  movel([-0.251057, -0.840337, -2.769867, -1.102185, 1.570796, 1.319739],accel_mss,speed_ms,0,blend_radius_m)
  movel([-0.250306, -0.839240, -2.770084, -1.103065, 1.570796, 1.320491],accel_mss,speed_ms,0,blend_radius_m)
  movel([-0.248421, -0.837227, -2.770480, -1.104681, 1.570796, 1.322375],accel_mss,speed_ms,0,blend_radius_m)
  movel([-0.247261, -0.836341, -2.770654, -1.105394, 1.570796, 1.323536],accel_mss,speed_ms,0,blend_radius_m)
  movel([-0.246051, -0.835788, -2.770763, -1.105839, 1.570796, 1.324746],accel_mss,speed_ms,0,blend_radius_m)
  movel([-0.245067, -0.835822, -2.770756, -1.105811, 1.570796, 1.325730],accel_mss,speed_ms,0,blend_radius_m)
  movel([-0.243698, -0.836942, -2.770537, -1.104911, 1.570796, 1.327098],accel_mss,speed_ms,0,blend_radius_m)
  movel([-0.242450, -0.839139, -2.770104, -1.103146, 1.570796, 1.328347],accel_mss,speed_ms,0,blend_radius_m)
  movel([-0.241508, -0.841625, -2.769611, -1.101153, 1.570796, 1.329288],accel_mss,speed_ms,0,blend_radius_m)
  movel([-0.239706, -0.837507, -2.770425, -1.104456, 1.570796, 1.331091],accel_mss,speed_ms,0,blend_radius_m)
  movel([-0.237551, -0.833302, -2.771247, -1.107840, 1.570796, 1.333246],accel_mss,speed_ms,0,blend_radius_m)
  movel([-0.235089, -0.829066, -2.772064, -1.111259, 1.570796, 1.335707],accel_mss,speed_ms,0,blend_radius_m)
  movel([-0.232380, -0.824862, -2.772866, -1.114661, 1.570796, 1.338416],accel_mss,speed_ms,0,blend_radius_m)
  movel([-0.226936, -0.816422, -2.774445, -1.121522, 1.570796, 1.343860],accel_mss,speed_ms,0,blend_radius_m)
  movel([-0.225279, -0.814079, -2.774877, -1.123434, 1.570796, 1.345517],accel_mss,speed_ms,0,blend_radius_m)
  movel([-0.223613, -0.811962, -2.775264, -1.125163, 1.570796, 1.347184],accel_mss,speed_ms,0,blend_radius_m)
  movel([-0.221984, -0.810225, -2.775580, -1.126584, 1.570796, 1.348813],accel_mss,speed_ms,0,blend_radius_m)
  movel([-0.220457, -0.809030, -2.775796, -1.127562, 1.570796, 1.350339],accel_mss,speed_ms,0,blend_radius_m)
  movel([-0.219063, -0.808558, -2.775882, -1.127949, 1.570796, 1.351734],accel_mss,speed_ms,0,blend_radius_m)
  movel([-0.217966, -0.808858, -2.775828, -1.127704, 1.570796, 1.352830],accel_mss,speed_ms,0,blend_radius_m)
  movel([-0.217165, -0.809769, -2.775663, -1.126958, 1.570796, 1.353632],accel_mss,speed_ms,0,blend_radius_m)
  movel([-0.216671, -0.811136, -2.775414, -1.125838, 1.570796, 1.354126],accel_mss,speed_ms,0,blend_radius_m)
  movel([-0.216485, -0.812799, -2.775111, -1.124479, 1.570796, 1.354311],accel_mss,speed_ms,0,blend_radius_m)
  movel([-0.216608, -0.814592, -2.774782, -1.123014, 1.570796, 1.354188],accel_mss,speed_ms,0,blend_radius_m)
  movel([-0.217044, -0.816361, -2.774456, -1.121571, 1.570796, 1.353752],accel_mss,speed_ms,0,blend_radius_m)
  movel([-0.217800, -0.817948, -2.774162, -1.120278, 1.570796, 1.352996],accel_mss,speed_ms,0,blend_radius_m)
  movel([-0.212688, -0.810429, -2.775543, -1.126417, 1.570796, 1.358108],accel_mss,speed_ms,0,blend_radius_m)
  movel([-0.209894, -0.806731, -2.776211, -1.129447, 1.570796, 1.360902],accel_mss,speed_ms,0,blend_radius_m)
  movel([-0.206949, -0.803115, -2.776856, -1.132417, 1.570796, 1.363847],accel_mss,speed_ms,0,blend_radius_m)
  movel([-0.203868, -0.799614, -2.777475, -1.135300, 1.570796, 1.366928],accel_mss,speed_ms,0,blend_radius_m)
  movel([-0.200656, -0.796258, -2.778062, -1.138069, 1.570796, 1.370141],accel_mss,speed_ms,0,blend_radius_m)
  movel([-0.197322, -0.793081, -2.778612, -1.140696, 1.570796, 1.373474],accel_mss,speed_ms,0,blend_radius_m)
  movel([-0.193879, -0.790113, -2.779121, -1.143155, 1.570796, 1.376917],accel_mss,speed_ms,0,blend_radius_m)
  movel([-0.191467, -0.788517, -2.779393, -1.144480, 1.570796, 1.379330],accel_mss,speed_ms,0,blend_radius_m)
  movel([-0.188786, -0.787373, -2.779587, -1.145430, 1.570796, 1.382010],accel_mss,speed_ms,0,blend_radius_m)
  movel([-0.187580, -0.787128, -2.779628, -1.145633, 1.570796, 1.383216],accel_mss,speed_ms,0,blend_radius_m)
  movel([-0.186584, -0.787179, -2.779619, -1.145591, 1.570796, 1.384213],accel_mss,speed_ms,0,blend_radius_m)
  movel([-0.185886, -0.787588, -2.779550, -1.145251, 1.570796, 1.384910],accel_mss,speed_ms,0,blend_radius_m)
  movel([-0.185586, -0.788421, -2.779409, -1.144559, 1.570796, 1.385210],accel_mss,speed_ms,0,blend_radius_m)
  movel([-0.185771, -0.789581, -2.779211, -1.143597, 1.570796, 1.385025],accel_mss,speed_ms,0,blend_radius_m)
  movel([-0.186325, -0.790924, -2.778982, -1.142483, 1.570796, 1.384471],accel_mss,speed_ms,0,blend_radius_m)
  movel([-0.188126, -0.794006, -2.778452, -1.139931, 1.570796, 1.382670],accel_mss,speed_ms,0,blend_radius_m)
  movel([-0.190402, -0.796962, -2.777939, -1.137488, 1.570796, 1.380394],accel_mss,speed_ms,0,blend_radius_m)
  movel([-0.192970, -0.799746, -2.777452, -1.135191, 1.570796, 1.377827],accel_mss,speed_ms,0,blend_radius_m)
  movel([-0.195646, -0.802312, -2.776999, -1.133078, 1.570796, 1.375151],accel_mss,speed_ms,0,blend_radius_m)
  movel([-0.191927, -0.800596, -2.777302, -1.134491, 1.570796, 1.378869],accel_mss,speed_ms,0,blend_radius_m)
  movel([-0.188109, -0.798487, -2.777673, -1.136229, 1.570796, 1.382688],accel_mss,speed_ms,0,blend_radius_m)
  movel([-0.184228, -0.796012, -2.778104, -1.138273, 1.570796, 1.386568],accel_mss,speed_ms,0,blend_radius_m)
  movel([-0.180320, -0.793191, -2.778593, -1.140606, 1.570796, 1.390476],accel_mss,speed_ms,0,blend_radius_m)
  movel([-0.177275, -0.790678, -2.779024, -1.142687, 1.570796, 1.393522],accel_mss,speed_ms,0,blend_radius_m)
  movel([-0.171365, -0.785323, -2.779933, -1.147134, 1.570796, 1.399431],accel_mss,speed_ms,0,blend_radius_m)
  movel([-0.168296, -0.782767, -2.780361, -1.149261, 1.570796, 1.402501],accel_mss,speed_ms,0,blend_radius_m)
  movel([-0.164758, -0.780078, -2.780808, -1.151503, 1.570796, 1.406038],accel_mss,speed_ms,0,blend_radius_m)
  movel([-0.158752, -0.775824, -2.781507, -1.155058, 1.570796, 1.412044],accel_mss,speed_ms,0,blend_radius_m)
  movel([-0.155841, -0.774007, -2.781803, -1.156579, 1.570796, 1.414955],accel_mss,speed_ms,0,blend_radius_m)
  movel([-0.153543, -0.772881, -2.781986, -1.157523, 1.570796, 1.417254],accel_mss,speed_ms,0,blend_radius_m)
  movel([-0.152751, -0.772687, -2.782017, -1.157685, 1.570796, 1.418046],accel_mss,speed_ms,0,blend_radius_m)
  movel([-0.152271, -0.772806, -2.781998, -1.157586, 1.570796, 1.418525],accel_mss,speed_ms,0,blend_radius_m)
  movel([-0.152148, -0.773270, -2.781923, -1.157196, 1.570796, 1.418648],accel_mss,speed_ms,0,blend_radius_m)
  movel([-0.152440, -0.774130, -2.781783, -1.156476, 1.570796, 1.418357],accel_mss,speed_ms,0,blend_radius_m)
  movel([-0.153723, -0.776356, -2.781420, -1.154613, 1.570796, 1.417074],accel_mss,speed_ms,0,blend_radius_m)
  movel([-0.155470, -0.778742, -2.781028, -1.152619, 1.570796, 1.415326],accel_mss,speed_ms,0,blend_radius_m)
  movel([-0.157553, -0.781219, -2.780619, -1.150552, 1.570796, 1.413244],accel_mss,speed_ms,0,blend_radius_m)
  movel([-0.159834, -0.783698, -2.780205, -1.148485, 1.570796, 1.410962],accel_mss,speed_ms,0,blend_radius_m)
  movel([-0.164497, -0.788374, -2.779417, -1.144598, 1.570796, 1.406299],accel_mss,speed_ms,0,blend_radius_m)
  movel([-0.168438, -0.792159, -2.778770, -1.141460, 1.570796, 1.402358],accel_mss,speed_ms,0,blend_radius_m)
  movel([-0.166238, -0.791550, -2.778875, -1.141964, 1.570796, 1.404559],accel_mss,speed_ms,0,blend_radius_m)
  movel([-0.163950, -0.790704, -2.779020, -1.142666, 1.570796, 1.406846],accel_mss,speed_ms,0,blend_radius_m)
  movel([-0.159176, -0.788425, -2.779408, -1.144556, 1.570796, 1.411620],accel_mss,speed_ms,0,blend_radius_m)
  movel([-0.154224, -0.785549, -2.779894, -1.146946, 1.570796, 1.416572],accel_mss,speed_ms,0,blend_radius_m)
  movel([-0.149200, -0.782306, -2.780438, -1.149645, 1.570796, 1.421597],accel_mss,speed_ms,0,blend_radius_m)
  movel([-0.145052, -0.779396, -2.780920, -1.152073, 1.570796, 1.425744],accel_mss,speed_ms,0,blend_radius_m)
  movel([-0.132523, -0.770152, -2.782425, -1.159811, 1.570796, 1.438273],accel_mss,speed_ms,0,blend_radius_m)
  movel([-0.130147, -0.768779, -2.782645, -1.160965, 1.570796, 1.440650],accel_mss,speed_ms,0,blend_radius_m)
  movel([-0.128213, -0.768174, -2.782742, -1.161473, 1.570796, 1.442583],accel_mss,speed_ms,0,blend_radius_m)
  movel([-0.127762, -0.768378, -2.782709, -1.161302, 1.570796, 1.443034],accel_mss,speed_ms,0,blend_radius_m)
  movel([-0.127842, -0.769035, -2.782604, -1.160750, 1.570796, 1.442955],accel_mss,speed_ms,0,blend_radius_m)
  movel([-0.128593, -0.770230, -2.782413, -1.159746, 1.570796, 1.442203],accel_mss,speed_ms,0,blend_radius_m)
  movel([-0.130154, -0.772048, -2.782120, -1.158221, 1.570796, 1.440642],accel_mss,speed_ms,0,blend_radius_m)
  movel([-0.132825, -0.774737, -2.781684, -1.155968, 1.570796, 1.437971],accel_mss,speed_ms,0,blend_radius_m)
  movel([-0.135952, -0.777548, -2.781225, -1.153616, 1.570796, 1.434844],accel_mss,speed_ms,0,blend_radius_m)
  movel([-0.139084, -0.779981, -2.780824, -1.151585, 1.570796, 1.431712],accel_mss,speed_ms,0,blend_radius_m)
  movel([-0.140515, -0.780901, -2.780671, -1.150816, 1.570796, 1.430281],accel_mss,speed_ms,0,blend_radius_m)
  movel([-0.141777, -0.781533, -2.780566, -1.150290, 1.570796, 1.429020],accel_mss,speed_ms,0,blend_radius_m)
  movel([-0.136604, -0.780701, -2.780705, -1.150984, 1.570796, 1.434192],accel_mss,speed_ms,0,blend_radius_m)
  movel([-0.131148, -0.779248, -2.780945, -1.152196, 1.570796, 1.439648],accel_mss,speed_ms,0,blend_radius_m)
  movel([-0.125468, -0.777292, -2.781267, -1.153830, 1.570796, 1.445329],accel_mss,speed_ms,0,blend_radius_m)
  movel([-0.119612, -0.774952, -2.781649, -1.155788, 1.570796, 1.451185],accel_mss,speed_ms,0,blend_radius_m)
  movel([-0.107622, -0.769590, -2.782515, -1.160284, 1.570796, 1.463175],accel_mss,speed_ms,0,blend_radius_m)
  movel([-0.095682, -0.764142, -2.783380, -1.164866, 1.570796, 1.475114],accel_mss,speed_ms,0,blend_radius_m)
  movel([-0.093660, -0.763518, -2.783479, -1.165393, 1.570796, 1.477136],accel_mss,speed_ms,0,blend_radius_m)
  movel([-0.092947, -0.763655, -2.783457, -1.165277, 1.570796, 1.477849],accel_mss,speed_ms,0,blend_radius_m)
  movel([-0.092662, -0.764296, -2.783356, -1.164736, 1.570796, 1.478134],accel_mss,speed_ms,0,blend_radius_m)
  movel([-0.092897, -0.765328, -2.783193, -1.163868, 1.570796, 1.477899],accel_mss,speed_ms,0,blend_radius_m)
  movel([-0.094551, -0.768317, -2.782719, -1.161353, 1.570796, 1.476245],accel_mss,speed_ms,0,blend_radius_m)
  movel([-0.095791, -0.770072, -2.782438, -1.159879, 1.570796, 1.475005],accel_mss,speed_ms,0,blend_radius_m)
  movel([-0.098671, -0.773409, -2.781900, -1.157080, 1.570796, 1.472125],accel_mss,speed_ms,0,blend_radius_m)
  movel([-0.101929, -0.776471, -2.781401, -1.154516, 1.570796, 1.468867],accel_mss,speed_ms,0,blend_radius_m)
  movel([-0.105410, -0.779237, -2.780947, -1.152206, 1.570796, 1.465387],accel_mss,speed_ms,0,blend_radius_m)
  movel([-0.108946, -0.781663, -2.780545, -1.150181, 1.570796, 1.461850],accel_mss,speed_ms,0,blend_radius_m)
  movel([-0.112381, -0.783724, -2.780201, -1.148464, 1.570796, 1.458416],accel_mss,speed_ms,0,blend_radius_m)
  movel([-0.115557, -0.785382, -2.779923, -1.147085, 1.570796, 1.455240],accel_mss,speed_ms,0,blend_radius_m)
  movel([-0.118308, -0.786594, -2.779718, -1.146077, 1.570796, 1.452489],accel_mss,speed_ms,0,blend_radius_m)
  movel([-0.118229, -0.787293, -2.779600, -1.145496, 1.570796, 1.452568],accel_mss,speed_ms,0,blend_radius_m)
  movel([-0.117672, -0.787561, -2.779555, -1.145274, 1.570796, 1.453124],accel_mss,speed_ms,0,blend_radius_m)
  movel([-0.116060, -0.787683, -2.779534, -1.145172, 1.570796, 1.454736],accel_mss,speed_ms,0,blend_radius_m)
  movel([-0.114280, -0.787508, -2.779564, -1.145318, 1.570796, 1.456517],accel_mss,speed_ms,0,blend_radius_m)
  movel([-0.110443, -0.786631, -2.779712, -1.146046, 1.570796, 1.460353],accel_mss,speed_ms,0,blend_radius_m)
  movel([-0.103651, -0.784713, -2.780035, -1.147641, 1.570796, 1.467145],accel_mss,speed_ms,0,blend_radius_m)
  movel([-0.096773, -0.782536, -2.780399, -1.149454, 1.570796, 1.474024],accel_mss,speed_ms,0,blend_radius_m)
  movel([-0.082734, -0.777500, -2.781233, -1.153657, 1.570796, 1.488063],accel_mss,speed_ms,0,blend_radius_m)
  movel([-0.078824, -0.776168, -2.781451, -1.154770, 1.570796, 1.491972],accel_mss,speed_ms,0,blend_radius_m)
  movel([-0.076323, -0.775517, -2.781557, -1.155315, 1.570796, 1.494474],accel_mss,speed_ms,0,blend_radius_m)
  movel([-0.073893, -0.775133, -2.781620, -1.155636, 1.570796, 1.496903],accel_mss,speed_ms,0,blend_radius_m)
  movel([-0.071878, -0.775218, -2.781606, -1.155565, 1.570796, 1.498918],accel_mss,speed_ms,0,blend_radius_m)
  movel([-0.070612, -0.775956, -2.781486, -1.154948, 1.570796, 1.500184],accel_mss,speed_ms,0,blend_radius_m)
  movel([-0.070357, -0.776623, -2.781377, -1.154390, 1.570796, 1.500439],accel_mss,speed_ms,0,blend_radius_m)
  movel([-0.070410, -0.777522, -2.781229, -1.153638, 1.570796, 1.500387],accel_mss,speed_ms,0,blend_radius_m)
  movel([-0.070817, -0.778683, -2.781038, -1.152668, 1.570796, 1.499979],accel_mss,speed_ms,0,blend_radius_m)
  movel([-0.071609, -0.780115, -2.780802, -1.151472, 1.570796, 1.499188],accel_mss,speed_ms,0,blend_radius_m)
  movel([-0.072883, -0.781500, -2.780572, -1.150317, 1.570796, 1.497913],accel_mss,speed_ms,0,blend_radius_m)
  movel([-0.074697, -0.782890, -2.780340, -1.149159, 1.570796, 1.496099],accel_mss,speed_ms,0,blend_radius_m)
  movel([-0.084551, -0.789376, -2.779246, -1.143767, 1.570796, 1.486245],accel_mss,speed_ms,0,blend_radius_m)
  movel([-0.087910, -0.791177, -2.778939, -1.142274, 1.570796, 1.482886],accel_mss,speed_ms,0,blend_radius_m)
  movel([-0.089384, -0.791747, -2.778841, -1.141801, 1.570796, 1.481412],accel_mss,speed_ms,0,blend_radius_m)
  movel([-0.090634, -0.791996, -2.778798, -1.141595, 1.570796, 1.480162],accel_mss,speed_ms,0,blend_radius_m)
  movel([-0.085187, -0.792592, -2.778696, -1.141101, 1.570796, 1.485610],accel_mss,speed_ms,0,blend_radius_m)
  movel([-0.079266, -0.792365, -2.778735, -1.141289, 1.570796, 1.491530],accel_mss,speed_ms,0,blend_radius_m)
  movel([-0.072987, -0.791466, -2.778889, -1.142034, 1.570796, 1.497810],accel_mss,speed_ms,0,blend_radius_m)
  movel([-0.066459, -0.790039, -2.779133, -1.143217, 1.570796, 1.504338],accel_mss,speed_ms,0,blend_radius_m)
  movel([-0.060916, -0.788133, -2.779458, -1.144799, 1.570796, 1.509880],accel_mss,speed_ms,0,blend_radius_m)
  movel([-0.052946, -0.785532, -2.779897, -1.146959, 1.570796, 1.517850],accel_mss,speed_ms,0,blend_radius_m)
  movel([-0.049278, -0.784724, -2.780033, -1.147631, 1.570796, 1.521518],accel_mss,speed_ms,0,blend_radius_m)
  movel([-0.046471, -0.784631, -2.780049, -1.147709, 1.570796, 1.524326],accel_mss,speed_ms,0,blend_radius_m)
  movel([-0.045545, -0.784943, -2.779996, -1.147450, 1.570796, 1.525252],accel_mss,speed_ms,0,blend_radius_m)
  movel([-0.045021, -0.785541, -2.779896, -1.146953, 1.570796, 1.525776],accel_mss,speed_ms,0,blend_radius_m)
  movel([-0.044956, -0.786463, -2.779740, -1.146186, 1.570796, 1.525840],accel_mss,speed_ms,0,blend_radius_m)
  movel([-0.045403, -0.787732, -2.779526, -1.145131, 1.570796, 1.525393],accel_mss,speed_ms,0,blend_radius_m)
  movel([-0.046180, -0.789074, -2.779298, -1.144017, 1.570796, 1.524616],accel_mss,speed_ms,0,blend_radius_m)
  movel([-0.047117, -0.790379, -2.779075, -1.142935, 1.570796, 1.523680],accel_mss,speed_ms,0,blend_radius_m)
  movel([-0.049250, -0.792857, -2.778650, -1.140882, 1.570796, 1.521546],accel_mss,speed_ms,0,blend_radius_m)
  movel([-0.051649, -0.795339, -2.778221, -1.138829, 1.570796, 1.519147],accel_mss,speed_ms,0,blend_radius_m)
  movel([-0.056596, -0.799831, -2.777437, -1.135121, 1.570796, 1.514200],accel_mss,speed_ms,0,blend_radius_m)
  movel([-0.059113, -0.801820, -2.777086, -1.133483, 1.570796, 1.511683],accel_mss,speed_ms,0,blend_radius_m)
  movel([-0.054139, -0.800667, -2.777290, -1.134433, 1.570796, 1.516658],accel_mss,speed_ms,0,blend_radius_m)
  movel([-0.049049, -0.799176, -2.777552, -1.135662, 1.570796, 1.521747],accel_mss,speed_ms,0,blend_radius_m)
  movel([-0.043853, -0.797385, -2.777865, -1.137138, 1.570796, 1.526944],accel_mss,speed_ms,0,blend_radius_m)
  movel([-0.038557, -0.795324, -2.778224, -1.138841, 1.570796, 1.532239],accel_mss,speed_ms,0,blend_radius_m)
  movel([-0.027716, -0.790540, -2.779048, -1.142802, 1.570796, 1.543080],accel_mss,speed_ms,0,blend_radius_m)
  movel([-0.016601, -0.785088, -2.779972, -1.147329, 1.570796, 1.554196],accel_mss,speed_ms,0,blend_radius_m)
  movel([-0.013645, -0.783918, -2.780168, -1.148302, 1.570796, 1.557151],accel_mss,speed_ms,0,blend_radius_m)
  movel([-0.012527, -0.783932, -2.780166, -1.148291, 1.570796, 1.558270],accel_mss,speed_ms,0,blend_radius_m)
  movel([-0.011960, -0.784664, -2.780043, -1.147681, 1.570796, 1.558836],accel_mss,speed_ms,0,blend_radius_m)
  movel([-0.011973, -0.785494, -2.779904, -1.146991, 1.570796, 1.558823],accel_mss,speed_ms,0,blend_radius_m)
  movel([-0.012257, -0.786461, -2.779741, -1.146187, 1.570796, 1.558540],accel_mss,speed_ms,0,blend_radius_m)
  movel([-0.013515, -0.788743, -2.779354, -1.144292, 1.570796, 1.557281],accel_mss,speed_ms,0,blend_radius_m)
  movel([-0.015472, -0.791310, -2.778916, -1.142163, 1.570796, 1.555324],accel_mss,speed_ms,0,blend_radius_m)
  movel([-0.017868, -0.793984, -2.778456, -1.139949, 1.570796, 1.552928],accel_mss,speed_ms,0,blend_radius_m)
  movel([-0.022942, -0.798903, -2.777600, -1.135886, 1.570796, 1.547854],accel_mss,speed_ms,0,blend_radius_m)
  movel([-0.026708, -0.802032, -2.777048, -1.133308, 1.570796, 1.544089],accel_mss,speed_ms,0,blend_radius_m)
  movel([-0.024456, -0.801160, -2.777202, -1.134026, 1.570796, 1.546340],accel_mss,speed_ms,0,blend_radius_m)
  movel([-0.022148, -0.800059, -2.777397, -1.134934, 1.570796, 1.548648],accel_mss,speed_ms,0,blend_radius_m)
  movel([-0.017405, -0.797244, -2.777890, -1.137255, 1.570796, 1.553391],accel_mss,speed_ms,0,blend_radius_m)
  movel([-0.012565, -0.793690, -2.778507, -1.140192, 1.570796, 1.558232],accel_mss,speed_ms,0,blend_radius_m)
  movel([-0.007710, -0.789520, -2.779222, -1.143648, 1.570796, 1.563087],accel_mss,speed_ms,0,blend_radius_m)
  movel([-0.002926, -0.784828, -2.780016, -1.147546, 1.570796, 1.567870],accel_mss,speed_ms,0,blend_radius_m)
  movel([0.001697, -0.779740, -2.780864, -1.151785, 1.570796, 1.572493],accel_mss,speed_ms,0,blend_radius_m)
  movel([0.006066, -0.774361, -2.781746, -1.156282, 1.570796, 1.576863],accel_mss,speed_ms,0,blend_radius_m)
  movel([0.010091, -0.768815, -2.782639, -1.160935, 1.570796, 1.580887],accel_mss,speed_ms,0,blend_radius_m)
  movel([0.011867, -0.766339, -2.783033, -1.163017, 1.570796, 1.582663],accel_mss,speed_ms,0,blend_radius_m)
  movel([0.012853, -0.765231, -2.783209, -1.163949, 1.570796, 1.583649],accel_mss,speed_ms,0,blend_radius_m)
  movel([0.013911, -0.764336, -2.783350, -1.164703, 1.570796, 1.584707],accel_mss,speed_ms,0,blend_radius_m)
  movel([0.015047, -0.763769, -2.783439, -1.165181, 1.570796, 1.585844],accel_mss,speed_ms,0,blend_radius_m)
  movel([0.016045, -0.763599, -2.783466, -1.165324, 1.570796, 1.586842],accel_mss,speed_ms,0,blend_radius_m)
  movel([0.017197, -0.764007, -2.783402, -1.164980, 1.570796, 1.587993],accel_mss,speed_ms,0,blend_radius_m)
  movel([0.017895, -0.765128, -2.783225, -1.164036, 1.570796, 1.588691],accel_mss,speed_ms,0,blend_radius_m)
  movel([0.018210, -0.766786, -2.782962, -1.162640, 1.570796, 1.589006],accel_mss,speed_ms,0,blend_radius_m)
  movel([0.018221, -0.768822, -2.782638, -1.160929, 1.570796, 1.589018],accel_mss,speed_ms,0,blend_radius_m)
  movel([0.017618, -0.773331, -2.781913, -1.157145, 1.570796, 1.588414],accel_mss,speed_ms,0,blend_radius_m)
  movel([0.016685, -0.777318, -2.781263, -1.153808, 1.570796, 1.587481],accel_mss,speed_ms,0,blend_radius_m)
  movel([0.020069, -0.771975, -2.782132, -1.158282, 1.570796, 1.590865],accel_mss,speed_ms,0,blend_radius_m)
  movel([0.023040, -0.766596, -2.782993, -1.162801, 1.570796, 1.593836],accel_mss,speed_ms,0,blend_radius_m)
  movel([0.025578, -0.761235, -2.783836, -1.167318, 1.570796, 1.596375],accel_mss,speed_ms,0,blend_radius_m)
  movel([0.027672, -0.755966, -2.784651, -1.171772, 1.570796, 1.598468],accel_mss,speed_ms,0,blend_radius_m)
  movel([0.029286, -0.750858, -2.785427, -1.176104, 1.570796, 1.600082],accel_mss,speed_ms,0,blend_radius_m)
  movel([0.030417, -0.745966, -2.786159, -1.180264, 1.570796, 1.601214],accel_mss,speed_ms,0,blend_radius_m)
  movel([0.031030, -0.741380, -2.786835, -1.184174, 1.570796, 1.601827],accel_mss,speed_ms,0,blend_radius_m)
  movel([0.031110, -0.737161, -2.787447, -1.187781, 1.570796, 1.601906],accel_mss,speed_ms,0,blend_radius_m)
  movel([0.030356, -0.731952, -2.788191, -1.192246, 1.570796, 1.601153],accel_mss,speed_ms,0,blend_radius_m)
  movel([0.030207, -0.729033, -2.788603, -1.194753, 1.570796, 1.601003],accel_mss,speed_ms,0,blend_radius_m)
  movel([0.030375, -0.727506, -2.788816, -1.196066, 1.570796, 1.601171],accel_mss,speed_ms,0,blend_radius_m)
  movel([0.030771, -0.725941, -2.789034, -1.197414, 1.570796, 1.601568],accel_mss,speed_ms,0,blend_radius_m)
  movel([0.031877, -0.723302, -2.789399, -1.199689, 1.570796, 1.602673],accel_mss,speed_ms,0,blend_radius_m)
  movel([0.033028, -0.721615, -2.789630, -1.201144, 1.570796, 1.603824],accel_mss,speed_ms,0,blend_radius_m)
  movel([0.034209, -0.720678, -2.789758, -1.201953, 1.570796, 1.605005],accel_mss,speed_ms,0,blend_radius_m)
  movel([0.035393, -0.720293, -2.789810, -1.202286, 1.570796, 1.606190],accel_mss,speed_ms,0,blend_radius_m)
  movel([0.038713, -0.720456, -2.789788, -1.202145, 1.570796, 1.609509],accel_mss,speed_ms,0,blend_radius_m)
  movel([0.039670, -0.720273, -2.789813, -1.202303, 1.570796, 1.610466],accel_mss,speed_ms,0,blend_radius_m)
  movel([0.041218, -0.716370, -2.790341, -1.205678, 1.570796, 1.612014],accel_mss,speed_ms,0,blend_radius_m)
  movel([0.042449, -0.712549, -2.790850, -1.208990, 1.570796, 1.613245],accel_mss,speed_ms,0,blend_radius_m)
  movel([0.043380, -0.708824, -2.791341, -1.212224, 1.570796, 1.614176],accel_mss,speed_ms,0,blend_radius_m)
  movel([0.044028, -0.705202, -2.791811, -1.215376, 1.570796, 1.614824],accel_mss,speed_ms,0,blend_radius_m)
  movel([0.044398, -0.701705, -2.792260, -1.218424, 1.570796, 1.615194],accel_mss,speed_ms,0,blend_radius_m)
  movel([0.044507, -0.698341, -2.792686, -1.221362, 1.570796, 1.615303],accel_mss,speed_ms,0,blend_radius_m)
  movel([0.044023, -0.692041, -2.793470, -1.226877, 1.570796, 1.614819],accel_mss,speed_ms,0,blend_radius_m)
  movel([0.042690, -0.686413, -2.794156, -1.231820, 1.570796, 1.613487],accel_mss,speed_ms,0,blend_radius_m)
  movel([0.040657, -0.681528, -2.794740, -1.236121, 1.570796, 1.611454],accel_mss,speed_ms,0,blend_radius_m)
  movel([0.038047, -0.677485, -2.795215, -1.239689, 1.570796, 1.608843],accel_mss,speed_ms,0,blend_radius_m)
  movel([0.035023, -0.674343, -2.795579, -1.242467, 1.570796, 1.605819],accel_mss,speed_ms,0,blend_radius_m)
  speed_ms = 0.005
  movel([0.035023, -0.668307, -2.788892, -1.255190, 1.570796, 1.605819],accel_mss,speed_ms,0,blend_radius_m)
  speed_ms = 0.040
  movel([0.005563, -0.693117, -2.785908, -1.233364, 1.570796, 1.576359],accel_mss,speed_ms,0,blend_radius_m)
  speed_ms = 0.005
  movel([0.005563, -0.699497, -2.792540, -1.220352, 1.570796, 1.576359],accel_mss,speed_ms,0,blend_radius_m)
  speed_ms = 0.025
  movel([0.002772, -0.699600, -2.792527, -1.220262, 1.570796, 1.573568],accel_mss,speed_ms,0,blend_radius_m)
  movel([-0.000362, -0.700496, -2.792414, -1.219480, 1.570796, 1.570434],accel_mss,speed_ms,0,blend_radius_m)
  movel([-0.003761, -0.702064, -2.792214, -1.218111, 1.570796, 1.567035],accel_mss,speed_ms,0,blend_radius_m)
  movel([-0.007341, -0.704171, -2.791944, -1.216274, 1.570796, 1.563455],accel_mss,speed_ms,0,blend_radius_m)
  movel([-0.011021, -0.706691, -2.791618, -1.214080, 1.570796, 1.559775],accel_mss,speed_ms,0,blend_radius_m)
  movel([-0.014730, -0.709498, -2.791252, -1.211639, 1.570796, 1.556067],accel_mss,speed_ms,0,blend_radius_m)
  movel([-0.021919, -0.715471, -2.790461, -1.206457, 1.570796, 1.548877],accel_mss,speed_ms,0,blend_radius_m)
  speed_ms = 0.005
  movel([-0.021919, -0.708883, -2.783866, -1.219640, 1.570796, 1.548877],accel_mss,speed_ms,0,blend_radius_m)
  speed_ms = 0.040
  movel([-0.012736, -0.700553, -2.784960, -1.226876, 1.570796, 1.558061],accel_mss,speed_ms,0,blend_radius_m)
  speed_ms = 0.005
  movel([-0.012736, -0.707032, -2.791574, -1.213783, 1.570796, 1.558061],accel_mss,speed_ms,0,blend_radius_m)
  speed_ms = 0.025
  movel([-0.011741, -0.702920, -2.792104, -1.217364, 1.570796, 1.559055],accel_mss,speed_ms,0,blend_radius_m)
  movel([-0.011148, -0.699151, -2.792584, -1.220654, 1.570796, 1.559648],accel_mss,speed_ms,0,blend_radius_m)
  movel([-0.010951, -0.695718, -2.793015, -1.223656, 1.570796, 1.559845],accel_mss,speed_ms,0,blend_radius_m)
  movel([-0.011133, -0.692605, -2.793401, -1.226383, 1.570796, 1.559663],accel_mss,speed_ms,0,blend_radius_m)
  movel([-0.011672, -0.689793, -2.793746, -1.228850, 1.570796, 1.559124],accel_mss,speed_ms,0,blend_radius_m)
  movel([-0.012556, -0.687267, -2.794053, -1.231069, 1.570796, 1.558241],accel_mss,speed_ms,0,blend_radius_m)
  movel([-0.013764, -0.685013, -2.794325, -1.233052, 1.570796, 1.557032],accel_mss,speed_ms,0,blend_radius_m)
  movel([-0.015280, -0.683011, -2.794564, -1.234815, 1.570796, 1.555516],accel_mss,speed_ms,0,blend_radius_m)
  movel([-0.020599, -0.678116, -2.795141, -1.239132, 1.570796, 1.550198],accel_mss,speed_ms,0,blend_radius_m)
  movel([-0.022981, -0.675592, -2.795435, -1.241363, 1.570796, 1.547815],accel_mss,speed_ms,0,blend_radius_m)
  movel([-0.024944, -0.672152, -2.795830, -1.244407, 1.570796, 1.545852],accel_mss,speed_ms,0,blend_radius_m)
  movel([-0.026696, -0.667138, -2.796398, -1.248853, 1.570796, 1.544100],accel_mss,speed_ms,0,blend_radius_m)
  movel([-0.027862, -0.661556, -2.797016, -1.253817, 1.570796, 1.542934],accel_mss,speed_ms,0,blend_radius_m)
  movel([-0.028220, -0.655275, -2.797696, -1.259418, 1.570796, 1.542576],accel_mss,speed_ms,0,blend_radius_m)
  movel([-0.028029, -0.651831, -2.798062, -1.262496, 1.570796, 1.542767],accel_mss,speed_ms,0,blend_radius_m)
  movel([-0.027547, -0.648162, -2.798446, -1.265781, 1.570796, 1.543250],accel_mss,speed_ms,0,blend_radius_m)
  movel([-0.026144, -0.642097, -2.799068, -1.271224, 1.570796, 1.544652],accel_mss,speed_ms,0,blend_radius_m)
  movel([-0.023952, -0.635758, -2.799701, -1.276930, 1.570796, 1.546845],accel_mss,speed_ms,0,blend_radius_m)
  movel([-0.020999, -0.629190, -2.800340, -1.282859, 1.570796, 1.549797],accel_mss,speed_ms,0,blend_radius_m)
  movel([-0.017318, -0.622446, -2.800977, -1.288965, 1.570796, 1.553478],accel_mss,speed_ms,0,blend_radius_m)
  movel([-0.012950, -0.615595, -2.801605, -1.295189, 1.570796, 1.557847],accel_mss,speed_ms,0,blend_radius_m)
  movel([-0.007925, -0.608692, -2.802219, -1.301478, 1.570796, 1.562872],accel_mss,speed_ms,0,blend_radius_m)
  movel([-0.002284, -0.601797, -2.802812, -1.307780, 1.570796, 1.568512],accel_mss,speed_ms,0,blend_radius_m)
  movel([0.003922, -0.594989, -2.803379, -1.314020, 1.570796, 1.574719],accel_mss,speed_ms,0,blend_radius_m)
  movel([0.008850, -0.590063, -2.803778, -1.318548, 1.570796, 1.579646],accel_mss,speed_ms,0,blend_radius_m)
  movel([0.013936, -0.585373, -2.804149, -1.322867, 1.570796, 1.584733],accel_mss,speed_ms,0,blend_radius_m)
  movel([0.019128, -0.580961, -2.804489, -1.326939, 1.570796, 1.589924],accel_mss,speed_ms,0,blend_radius_m)
  movel([0.024383, -0.576845, -2.804800, -1.330743, 1.570796, 1.595179],accel_mss,speed_ms,0,blend_radius_m)
  movel([0.029644, -0.573079, -2.805079, -1.334231, 1.570796, 1.600440],accel_mss,speed_ms,0,blend_radius_m)
  movel([0.034862, -0.569690, -2.805325, -1.337374, 1.570796, 1.605658],accel_mss,speed_ms,0,blend_radius_m)
  movel([0.039979, -0.566716, -2.805537, -1.340135, 1.570796, 1.610775],accel_mss,speed_ms,0,blend_radius_m)
  movel([0.044944, -0.564196, -2.805715, -1.342479, 1.570796, 1.615740],accel_mss,speed_ms,0,blend_radius_m)
  movel([0.049699, -0.562164, -2.805856, -1.344369, 1.570796, 1.620495],accel_mss,speed_ms,0,blend_radius_m)
  movel([0.054199, -0.560647, -2.805960, -1.345782, 1.570796, 1.624995],accel_mss,speed_ms,0,blend_radius_m)
  movel([0.058387, -0.559683, -2.806026, -1.346680, 1.570796, 1.629184],accel_mss,speed_ms,0,blend_radius_m)
  movel([0.062215, -0.559301, -2.806052, -1.347036, 1.570796, 1.633011],accel_mss,speed_ms,0,blend_radius_m)
  movel([0.065633, -0.559525, -2.806036, -1.346827, 1.570796, 1.636430],accel_mss,speed_ms,0,blend_radius_m)
  movel([0.068583, -0.560396, -2.805977, -1.346016, 1.570796, 1.639379],accel_mss,speed_ms,0,blend_radius_m)
  movel([0.071026, -0.561923, -2.805872, -1.344593, 1.570796, 1.641822],accel_mss,speed_ms,0,blend_radius_m)
  movel([0.072920, -0.564138, -2.805719, -1.342532, 1.570796, 1.643716],accel_mss,speed_ms,0,blend_radius_m)
  movel([0.074676, -0.567785, -2.805462, -1.339142, 1.570796, 1.645473],accel_mss,speed_ms,0,blend_radius_m)
  movel([0.075891, -0.571973, -2.805160, -1.335256, 1.570796, 1.646687],accel_mss,speed_ms,0,blend_radius_m)
  movel([0.076668, -0.576581, -2.804820, -1.330988, 1.570796, 1.647464],accel_mss,speed_ms,0,blend_radius_m)
  movel([0.077130, -0.581463, -2.804451, -1.326475, 1.570796, 1.647927],accel_mss,speed_ms,0,blend_radius_m)
  movel([0.077482, -0.592588, -2.803575, -1.316226, 1.570796, 1.648279],accel_mss,speed_ms,0,blend_radius_m)
  movel([0.077191, -0.604219, -2.802606, -1.305564, 1.570796, 1.647987],accel_mss,speed_ms,0,blend_radius_m)
  movel([0.076408, -0.616212, -2.801550, -1.294627, 1.570796, 1.647204],accel_mss,speed_ms,0,blend_radius_m)
  movel([0.075281, -0.628414, -2.800414, -1.283560, 1.570796, 1.646077],accel_mss,speed_ms,0,blend_radius_m)
  movel([0.070103, -0.676768, -2.795298, -1.240323, 1.570796, 1.640899],accel_mss,speed_ms,0,blend_radius_m)
  movel([0.068408, -0.699650, -2.792521, -1.220218, 1.570796, 1.639204],accel_mss,speed_ms,0,blend_radius_m)
  movel([0.067946, -0.710698, -2.791095, -1.210596, 1.570796, 1.638742],accel_mss,speed_ms,0,blend_radius_m)
  movel([0.067855, -0.721372, -2.789663, -1.201354, 1.570796, 1.638651],accel_mss,speed_ms,0,blend_radius_m)
  movel([0.068210, -0.731613, -2.788239, -1.192537, 1.570796, 1.639006],accel_mss,speed_ms,0,blend_radius_m)
  movel([0.069087, -0.741348, -2.786839, -1.184202, 1.570796, 1.639884],accel_mss,speed_ms,0,blend_radius_m)
  movel([0.070552, -0.750526, -2.785477, -1.176385, 1.570796, 1.641348],accel_mss,speed_ms,0,blend_radius_m)
  movel([0.072685, -0.759083, -2.784170, -1.169135, 1.570796, 1.643482],accel_mss,speed_ms,0,blend_radius_m)
  movel([0.073786, -0.762163, -2.783691, -1.166535, 1.570796, 1.644583],accel_mss,speed_ms,0,blend_radius_m)
  movel([0.075340, -0.764775, -2.783281, -1.164333, 1.570796, 1.646136],accel_mss,speed_ms,0,blend_radius_m)
  movel([0.077562, -0.766509, -2.783007, -1.162874, 1.570796, 1.648359],accel_mss,speed_ms,0,blend_radius_m)
  movel([0.078995, -0.766915, -2.782942, -1.162532, 1.570796, 1.649791],accel_mss,speed_ms,0,blend_radius_m)
  movel([0.080684, -0.766942, -2.782938, -1.162510, 1.570796, 1.651480],accel_mss,speed_ms,0,blend_radius_m)
  speed_ms = 0.005
  movel([0.080684, -0.759735, -2.776473, -1.176181, 1.570796, 1.651480],accel_mss,speed_ms,0,blend_radius_m)
  speed_ms = 0.040
  movel([0.042306, -0.732546, -2.780582, -1.199261, 1.570796, 1.613102],accel_mss,speed_ms,0,blend_radius_m)
  speed_ms = 0.005
  movel([0.042306, -0.739433, -2.787118, -1.185838, 1.570796, 1.613102],accel_mss,speed_ms,0,blend_radius_m)
  speed_ms = 0.025
  movel([0.041280, -0.741224, -2.786857, -1.184307, 1.570796, 1.612077],accel_mss,speed_ms,0,blend_radius_m)
  movel([0.040567, -0.743006, -2.786596, -1.182786, 1.570796, 1.611363],accel_mss,speed_ms,0,blend_radius_m)
  movel([0.040141, -0.744758, -2.786338, -1.181293, 1.570796, 1.610937],accel_mss,speed_ms,0,blend_radius_m)
  movel([0.039950, -0.746497, -2.786080, -1.179811, 1.570796, 1.610746],accel_mss,speed_ms,0,blend_radius_m)
  movel([0.040162, -0.749894, -2.785573, -1.176922, 1.570796, 1.610958],accel_mss,speed_ms,0,blend_radius_m)
  movel([0.040914, -0.753176, -2.785076, -1.174136, 1.570796, 1.611710],accel_mss,speed_ms,0,blend_radius_m)
  movel([0.043645, -0.762084, -2.783703, -1.166602, 1.570796, 1.614441],accel_mss,speed_ms,0,blend_radius_m)
  movel([0.043802, -0.764642, -2.783302, -1.164445, 1.570796, 1.614598],accel_mss,speed_ms,0,blend_radius_m)
  movel([0.043451, -0.765976, -2.783091, -1.163322, 1.570796, 1.614248],accel_mss,speed_ms,0,blend_radius_m)
  movel([0.042681, -0.767183, -2.782899, -1.162307, 1.570796, 1.613477],accel_mss,speed_ms,0,blend_radius_m)
  movel([0.041894, -0.767952, -2.782777, -1.161660, 1.570796, 1.612690],accel_mss,speed_ms,0,blend_radius_m)
  movel([0.041097, -0.768332, -2.782717, -1.161341, 1.570796, 1.611893],accel_mss,speed_ms,0,blend_radius_m)
  movel([0.040296, -0.768377, -2.782709, -1.161302, 1.570796, 1.611092],accel_mss,speed_ms,0,blend_radius_m)
  movel([0.038725, -0.767634, -2.782828, -1.161927, 1.570796, 1.609521],accel_mss,speed_ms,0,blend_radius_m)
  movel([0.037253, -0.766108, -2.783070, -1.163211, 1.570796, 1.608050],accel_mss,speed_ms,0,blend_radius_m)
  movel([0.034904, -0.762212, -2.783683, -1.166494, 1.570796, 1.605700],accel_mss,speed_ms,0,blend_radius_m)
  movel([0.033908, -0.759677, -2.784078, -1.168634, 1.570796, 1.604705],accel_mss,speed_ms,0,blend_radius_m)
  movel([0.032880, -0.764620, -2.783305, -1.164464, 1.570796, 1.603677],accel_mss,speed_ms,0,blend_radius_m)
  movel([0.032537, -0.769144, -2.782587, -1.160658, 1.570796, 1.603333],accel_mss,speed_ms,0,blend_radius_m)
  movel([0.032771, -0.773293, -2.781919, -1.157177, 1.570796, 1.603568],accel_mss,speed_ms,0,blend_radius_m)
  movel([0.033490, -0.777081, -2.781301, -1.154007, 1.570796, 1.604286],accel_mss,speed_ms,0,blend_radius_m)
  movel([0.034586, -0.780554, -2.780729, -1.151106, 1.570796, 1.605382],accel_mss,speed_ms,0,blend_radius_m)
  movel([0.035975, -0.783720, -2.780202, -1.148468, 1.570796, 1.606771],accel_mss,speed_ms,0,blend_radius_m)
  movel([0.039232, -0.789251, -2.779268, -1.143870, 1.570796, 1.610029],accel_mss,speed_ms,0,blend_radius_m)
  movel([0.039501, -0.790641, -2.779031, -1.142718, 1.570796, 1.610298],accel_mss,speed_ms,0,blend_radius_m)
  movel([0.039228, -0.791488, -2.778885, -1.142015, 1.570796, 1.610024],accel_mss,speed_ms,0,blend_radius_m)
  movel([0.038582, -0.792263, -2.778752, -1.141373, 1.570796, 1.609379],accel_mss,speed_ms,0,blend_radius_m)
  movel([0.037678, -0.792716, -2.778675, -1.140998, 1.570796, 1.608474],accel_mss,speed_ms,0,blend_radius_m)
  movel([0.035647, -0.793134, -2.778603, -1.140653, 1.570796, 1.606443],accel_mss,speed_ms,0,blend_radius_m)
  movel([0.033888, -0.793076, -2.778612, -1.140700, 1.570796, 1.604685],accel_mss,speed_ms,0,blend_radius_m)
  movel([0.032370, -0.792615, -2.778692, -1.141082, 1.570796, 1.603166],accel_mss,speed_ms,0,blend_radius_m)
  movel([0.031075, -0.791799, -2.778832, -1.141758, 1.570796, 1.601871],accel_mss,speed_ms,0,blend_radius_m)
  movel([0.029067, -0.789360, -2.779249, -1.143780, 1.570796, 1.599863],accel_mss,speed_ms,0,blend_radius_m)
  movel([0.027691, -0.786242, -2.779778, -1.146369, 1.570796, 1.598487],accel_mss,speed_ms,0,blend_radius_m)
  movel([0.028004, -0.793796, -2.778488, -1.140105, 1.570796, 1.598800],accel_mss,speed_ms,0,blend_radius_m)
  movel([0.028562, -0.797205, -2.777897, -1.137288, 1.570796, 1.599358],accel_mss,speed_ms,0,blend_radius_m)
  movel([0.029625, -0.800190, -2.777373, -1.134825, 1.570796, 1.600421],accel_mss,speed_ms,0,blend_radius_m)
  movel([0.031179, -0.802173, -2.777023, -1.133193, 1.570796, 1.601975],accel_mss,speed_ms,0,blend_radius_m)
  movel([0.034992, -0.805024, -2.776516, -1.130849, 1.570796, 1.605788],accel_mss,speed_ms,0,blend_radius_m)
  movel([0.036442, -0.807008, -2.776161, -1.129220, 1.570796, 1.607238],accel_mss,speed_ms,0,blend_radius_m)
  movel([0.036608, -0.807530, -2.776067, -1.128792, 1.570796, 1.607404],accel_mss,speed_ms,0,blend_radius_m)
  movel([0.036507, -0.808227, -2.775941, -1.128220, 1.570796, 1.607303],accel_mss,speed_ms,0,blend_radius_m)
  movel([0.035964, -0.809029, -2.775797, -1.127563, 1.570796, 1.606760],accel_mss,speed_ms,0,blend_radius_m)
  movel([0.034988, -0.809856, -2.775647, -1.126886, 1.570796, 1.605784],accel_mss,speed_ms,0,blend_radius_m)
  movel([0.032292, -0.811462, -2.775355, -1.125572, 1.570796, 1.603088],accel_mss,speed_ms,0,blend_radius_m)
  movel([0.027761, -0.813504, -2.774982, -1.123903, 1.570796, 1.598557],accel_mss,speed_ms,0,blend_radius_m)
  movel([0.028593, -0.815315, -2.774649, -1.122425, 1.570796, 1.599390],accel_mss,speed_ms,0,blend_radius_m)
  movel([0.029787, -0.817216, -2.774298, -1.120875, 1.570796, 1.600583],accel_mss,speed_ms,0,blend_radius_m)
  movel([0.031420, -0.819047, -2.773958, -1.119384, 1.570796, 1.602216],accel_mss,speed_ms,0,blend_radius_m)
  movel([0.033576, -0.820652, -2.773659, -1.118079, 1.570796, 1.604372],accel_mss,speed_ms,0,blend_radius_m)
  movel([0.039438, -0.821730, -2.773457, -1.117203, 1.570796, 1.610235],accel_mss,speed_ms,0,blend_radius_m)
  movel([0.042687, -0.822474, -2.773317, -1.116598, 1.570796, 1.613483],accel_mss,speed_ms,0,blend_radius_m)
  movel([0.043646, -0.822972, -2.773223, -1.116194, 1.570796, 1.614443],accel_mss,speed_ms,0,blend_radius_m)
  movel([0.043885, -0.823578, -2.773109, -1.115702, 1.570796, 1.614681],accel_mss,speed_ms,0,blend_radius_m)
  movel([0.043526, -0.824377, -2.772958, -1.115054, 1.570796, 1.614322],accel_mss,speed_ms,0,blend_radius_m)
  movel([0.042958, -0.825169, -2.772808, -1.114413, 1.570796, 1.613754],accel_mss,speed_ms,0,blend_radius_m)
  movel([0.041525, -0.826462, -2.772562, -1.113365, 1.570796, 1.612322],accel_mss,speed_ms,0,blend_radius_m)
  movel([0.040307, -0.827109, -2.772439, -1.112842, 1.570796, 1.611103],accel_mss,speed_ms,0,blend_radius_m)
  movel([0.039076, -0.827542, -2.772356, -1.112491, 1.570796, 1.609872],accel_mss,speed_ms,0,blend_radius_m)
  movel([0.036734, -0.828192, -2.772232, -1.111965, 1.570796, 1.607530],accel_mss,speed_ms,0,blend_radius_m)
  movel([0.037952, -0.830627, -2.771764, -1.109998, 1.570796, 1.608749],accel_mss,speed_ms,0,blend_radius_m)
  movel([0.039422, -0.832797, -2.771345, -1.108247, 1.570796, 1.610219],accel_mss,speed_ms,0,blend_radius_m)
  movel([0.041139, -0.834692, -2.770977, -1.106721, 1.570796, 1.611936],accel_mss,speed_ms,0,blend_radius_m)
  movel([0.043079, -0.836318, -2.770659, -1.105412, 1.570796, 1.613876],accel_mss,speed_ms,0,blend_radius_m)
  movel([0.045345, -0.837473, -2.770432, -1.104484, 1.570796, 1.616141],accel_mss,speed_ms,0,blend_radius_m)
  movel([0.047969, -0.838110, -2.770307, -1.103972, 1.570796, 1.618765],accel_mss,speed_ms,0,blend_radius_m)
  movel([0.053679, -0.838640, -2.770202, -1.103546, 1.570796, 1.624476],accel_mss,speed_ms,0,blend_radius_m)
  movel([0.055146, -0.839101, -2.770111, -1.103177, 1.570796, 1.625942],accel_mss,speed_ms,0,blend_radius_m)
  movel([0.055501, -0.839710, -2.769991, -1.102688, 1.570796, 1.626297],accel_mss,speed_ms,0,blend_radius_m)
  movel([0.055369, -0.840676, -2.769800, -1.101914, 1.570796, 1.626165],accel_mss,speed_ms,0,blend_radius_m)
  movel([0.054832, -0.841662, -2.769604, -1.101123, 1.570796, 1.625629],accel_mss,speed_ms,0,blend_radius_m)
  movel([0.054049, -0.842575, -2.769422, -1.100392, 1.570796, 1.624846],accel_mss,speed_ms,0,blend_radius_m)
  movel([0.052179, -0.844093, -2.769119, -1.099177, 1.570796, 1.622976],accel_mss,speed_ms,0,blend_radius_m)
  movel([0.049682, -0.845645, -2.768807, -1.097937, 1.570796, 1.620478],accel_mss,speed_ms,0,blend_radius_m)
  movel([0.047262, -0.846874, -2.768559, -1.096955, 1.570796, 1.618058],accel_mss,speed_ms,0,blend_radius_m)
  movel([0.044909, -0.847832, -2.768366, -1.096191, 1.570796, 1.615705],accel_mss,speed_ms,0,blend_radius_m)
  movel([0.042620, -0.848549, -2.768220, -1.095620, 1.570796, 1.613417],accel_mss,speed_ms,0,blend_radius_m)
  movel([0.044189, -0.850146, -2.767896, -1.094348, 1.570796, 1.614986],accel_mss,speed_ms,0,blend_radius_m)
  movel([0.046037, -0.851375, -2.767645, -1.093369, 1.570796, 1.616834],accel_mss,speed_ms,0,blend_radius_m)
  movel([0.048153, -0.852198, -2.767476, -1.092715, 1.570796, 1.618950],accel_mss,speed_ms,0,blend_radius_m)
  movel([0.050527, -0.852584, -2.767397, -1.092408, 1.570796, 1.621323],accel_mss,speed_ms,0,blend_radius_m)
  movel([0.053159, -0.852492, -2.767416, -1.092481, 1.570796, 1.623955],accel_mss,speed_ms,0,blend_radius_m)
  movel([0.056044, -0.851886, -2.767540, -1.092962, 1.570796, 1.626840],accel_mss,speed_ms,0,blend_radius_m)
  movel([0.059177, -0.850724, -2.767778, -1.093887, 1.570796, 1.629974],accel_mss,speed_ms,0,blend_radius_m)
  movel([0.062561, -0.848967, -2.768136, -1.095287, 1.570796, 1.633358],accel_mss,speed_ms,0,blend_radius_m)
  speed_ms = 0.005
  movel([0.062561, -0.840951, -2.761912, -1.109527, 1.570796, 1.633358],accel_mss,speed_ms,0,blend_radius_m)
  speed_ms = 0.040
  movel([0.075795, -0.818881, -2.766224, -1.127284, 1.570796, 1.646591],accel_mss,speed_ms,0,blend_radius_m)
  speed_ms = 0.005
  movel([0.075795, -0.826699, -2.772517, -1.113173, 1.570796, 1.646591],accel_mss,speed_ms,0,blend_radius_m)
  speed_ms = 0.025
  movel([0.069246, -0.827412, -2.772381, -1.112596, 1.570796, 1.640042],accel_mss,speed_ms,0,blend_radius_m)
  movel([0.066435, -0.827449, -2.772374, -1.112566, 1.570796, 1.637231],accel_mss,speed_ms,0,blend_radius_m)
  movel([0.063902, -0.827186, -2.772424, -1.112779, 1.570796, 1.634698],accel_mss,speed_ms,0,blend_radius_m)
  movel([0.061616, -0.826556, -2.772544, -1.113289, 1.570796, 1.632412],accel_mss,speed_ms,0,blend_radius_m)
  movel([0.059553, -0.825496, -2.772746, -1.114148, 1.570796, 1.630350],accel_mss,speed_ms,0,blend_radius_m)
  movel([0.057681, -0.823946, -2.773039, -1.115404, 1.570796, 1.628477],accel_mss,speed_ms,0,blend_radius_m)
  movel([0.055980, -0.821837, -2.773436, -1.117116, 1.570796, 1.626776],accel_mss,speed_ms,0,blend_radius_m)
  movel([0.053108, -0.816711, -2.774392, -1.121286, 1.570796, 1.623905],accel_mss,speed_ms,0,blend_radius_m)
  movel([0.050882, -0.810920, -2.775454, -1.126015, 1.570796, 1.621678],accel_mss,speed_ms,0,blend_radius_m)
  movel([0.049243, -0.804547, -2.776601, -1.131241, 1.570796, 1.620039],accel_mss,speed_ms,0,blend_radius_m)
  movel([0.048128, -0.797692, -2.777812, -1.136885, 1.570796, 1.618924],accel_mss,speed_ms,0,blend_radius_m)
  movel([0.047601, -0.791744, -2.778841, -1.141803, 1.570796, 1.618397],accel_mss,speed_ms,0,blend_radius_m)
  movel([0.047385, -0.785532, -2.779897, -1.146960, 1.570796, 1.618182],accel_mss,speed_ms,0,blend_radius_m)
  movel([0.047646, -0.772473, -2.782052, -1.157865, 1.570796, 1.618442],accel_mss,speed_ms,0,blend_radius_m)
  movel([0.049995, -0.725660, -2.789073, -1.197656, 1.570796, 1.620792],accel_mss,speed_ms,0,blend_radius_m)
  movel([0.050399, -0.715701, -2.790430, -1.206258, 1.570796, 1.621195],accel_mss,speed_ms,0,blend_radius_m)
  movel([0.050580, -0.705827, -2.791730, -1.214832, 1.570796, 1.621376],accel_mss,speed_ms,0,blend_radius_m)
  movel([0.050384, -0.696205, -2.792954, -1.223230, 1.570796, 1.621180],accel_mss,speed_ms,0,blend_radius_m)
  movel([0.049644, -0.687000, -2.794085, -1.231303, 1.570796, 1.620440],accel_mss,speed_ms,0,blend_radius_m)
  movel([0.048197, -0.678390, -2.795109, -1.238890, 1.570796, 1.618994],accel_mss,speed_ms,0,blend_radius_m)
  movel([0.045872, -0.670562, -2.796011, -1.245815, 1.570796, 1.616668],accel_mss,speed_ms,0,blend_radius_m)
  movel([0.043563, -0.665435, -2.796588, -1.250367, 1.570796, 1.614360],accel_mss,speed_ms,0,blend_radius_m)
  movel([0.040666, -0.660693, -2.797111, -1.254586, 1.570796, 1.611462],accel_mss,speed_ms,0,blend_radius_m)
  movel([0.037156, -0.656487, -2.797566, -1.258336, 1.570796, 1.607953],accel_mss,speed_ms,0,blend_radius_m)
  movel([0.033011, -0.652965, -2.797942, -1.261482, 1.570796, 1.603807],accel_mss,speed_ms,0,blend_radius_m)
  movel([0.028220, -0.650266, -2.798226, -1.263896, 1.570796, 1.599016],accel_mss,speed_ms,0,blend_radius_m)
  movel([0.022773, -0.648525, -2.798408, -1.265456, 1.570796, 1.593570],accel_mss,speed_ms,0,blend_radius_m)
  movel([0.016661, -0.647891, -2.798474, -1.266024, 1.570796, 1.587458],accel_mss,speed_ms,0,blend_radius_m)
  movel([0.009900, -0.648482, -2.798413, -1.265495, 1.570796, 1.580696],accel_mss,speed_ms,0,blend_radius_m)
  movel([0.006477, -0.649269, -2.798331, -1.264790, 1.570796, 1.577273],accel_mss,speed_ms,0,blend_radius_m)
  movel([0.002850, -0.650460, -2.798206, -1.263723, 1.570796, 1.573646],accel_mss,speed_ms,0,blend_radius_m)
  movel([-0.000948, -0.652066, -2.798037, -1.262286, 1.570796, 1.569848],accel_mss,speed_ms,0,blend_radius_m)
  movel([-0.004873, -0.654090, -2.797823, -1.260477, 1.570796, 1.565924],accel_mss,speed_ms,0,blend_radius_m)
  movel([-0.008880, -0.656522, -2.797563, -1.258305, 1.570796, 1.561917],accel_mss,speed_ms,0,blend_radius_m)
  movel([-0.012939, -0.659379, -2.797254, -1.255756, 1.570796, 1.557857],accel_mss,speed_ms,0,blend_radius_m)
  movel([-0.017001, -0.662646, -2.796896, -1.252847, 1.570796, 1.553795],accel_mss,speed_ms,0,blend_radius_m)
  movel([-0.021024, -0.666329, -2.796488, -1.249572, 1.570796, 1.549772],accel_mss,speed_ms,0,blend_radius_m)
  speed_ms = 0.005
  movel([-0.021024, -0.660405, -2.789785, -1.262198, 1.570796, 1.549772],accel_mss,speed_ms,0,blend_radius_m)
  speed_ms = 0.040
  movel([-0.038128, -0.652576, -2.790643, -1.269170, 1.570796, 1.532668],accel_mss,speed_ms,0,blend_radius_m)
  speed_ms = 0.005
  movel([-0.038128, -0.658385, -2.797362, -1.256642, 1.570796, 1.532668],accel_mss,speed_ms,0,blend_radius_m)
  speed_ms = 0.025
  movel([-0.038997, -0.656585, -2.797556, -1.258248, 1.570796, 1.531800],accel_mss,speed_ms,0,blend_radius_m)
  movel([-0.039545, -0.654488, -2.797780, -1.260121, 1.570796, 1.531251],accel_mss,speed_ms,0,blend_radius_m)
  movel([-0.039863, -0.649596, -2.798296, -1.264496, 1.570796, 1.530934],accel_mss,speed_ms,0,blend_radius_m)
  movel([-0.039428, -0.644050, -2.798869, -1.269470, 1.570796, 1.531368],accel_mss,speed_ms,0,blend_radius_m)
  movel([-0.038606, -0.638221, -2.799457, -1.274711, 1.570796, 1.532190],accel_mss,speed_ms,0,blend_radius_m)
  speed_ms = 0.005
  movel([-0.038606, -0.632709, -2.792700, -1.286981, 1.570796, 1.532190],accel_mss,speed_ms,0,blend_radius_m)
  speed_ms = 0.040
  movel([-0.029244, -0.628573, -2.793107, -1.290709, 1.570796, 1.541552],accel_mss,speed_ms,0,blend_radius_m)
  speed_ms = 0.005
  movel([-0.029244, -0.634022, -2.799872, -1.278495, 1.570796, 1.541552],accel_mss,speed_ms,0,blend_radius_m)
  speed_ms = 0.025
  movel([-0.030726, -0.633100, -2.799962, -1.279326, 1.570796, 1.540071],accel_mss,speed_ms,0,blend_radius_m)
  movel([-0.031885, -0.631872, -2.800082, -1.280435, 1.570796, 1.538911],accel_mss,speed_ms,0,blend_radius_m)
  movel([-0.033329, -0.628578, -2.800399, -1.283412, 1.570796, 1.537467],accel_mss,speed_ms,0,blend_radius_m)
  movel([-0.033718, -0.624318, -2.800802, -1.287269, 1.570796, 1.537078],accel_mss,speed_ms,0,blend_radius_m)
  movel([-0.033197, -0.619259, -2.801272, -1.291858, 1.570796, 1.537599],accel_mss,speed_ms,0,blend_radius_m)
  movel([-0.031911, -0.613583, -2.801786, -1.297020, 1.570796, 1.538885],accel_mss,speed_ms,0,blend_radius_m)
  movel([-0.030009, -0.607474, -2.802325, -1.302590, 1.570796, 1.540788],accel_mss,speed_ms,0,blend_radius_m)
  movel([-0.027642, -0.601117, -2.802870, -1.308402, 1.570796, 1.543154],accel_mss,speed_ms,0,blend_radius_m)
  movel([-0.024970, -0.594710, -2.803402, -1.314277, 1.570796, 1.545826],accel_mss,speed_ms,0,blend_radius_m)
  speed_ms = 0.005
  movel([-0.024970, -0.589875, -2.796570, -1.325944, 1.570796, 1.545826],accel_mss,speed_ms,0,blend_radius_m)
  speed_ms = 0.040
  movel([0.014719, -0.527887, -2.800866, -1.383636, 1.570796, 1.585515],accel_mss,speed_ms,0,blend_radius_m)
  speed_ms = 0.005
  movel([0.014719, -0.531662, -2.807783, -1.372944, 1.570796, 1.585515],accel_mss,speed_ms,0,blend_radius_m)
  speed_ms = 0.025
  movel([0.010416, -0.537007, -2.807471, -1.367911, 1.570796, 1.581212],accel_mss,speed_ms,0,blend_radius_m)
  movel([0.006202, -0.542586, -2.807133, -1.362670, 1.570796, 1.576999],accel_mss,speed_ms,0,blend_radius_m)
  movel([0.002146, -0.548310, -2.806775, -1.357304, 1.570796, 1.572943],accel_mss,speed_ms,0,blend_radius_m)
  movel([-0.001706, -0.554114, -2.806399, -1.351876, 1.570796, 1.569090],accel_mss,speed_ms,0,blend_radius_m)
  movel([-0.005287, -0.559918, -2.806010, -1.346461, 1.570796, 1.565509],accel_mss,speed_ms,0,blend_radius_m)
  movel([-0.008550, -0.565646, -2.805613, -1.341130, 1.570796, 1.562247],accel_mss,speed_ms,0,blend_radius_m)
  movel([-0.011435, -0.571233, -2.805214, -1.335943, 1.570796, 1.559361],accel_mss,speed_ms,0,blend_radius_m)
  movel([-0.013894, -0.576610, -2.804818, -1.330961, 1.570796, 1.556902],accel_mss,speed_ms,0,blend_radius_m)
  movel([-0.015880, -0.581704, -2.804433, -1.326252, 1.570796, 1.554916],accel_mss,speed_ms,0,blend_radius_m)
  movel([-0.017347, -0.586460, -2.804064, -1.321865, 1.570796, 1.553450],accel_mss,speed_ms,0,blend_radius_m)
  movel([-0.018248, -0.590811, -2.803718, -1.317860, 1.570796, 1.552549],accel_mss,speed_ms,0,blend_radius_m)
  movel([-0.018539, -0.594697, -2.803403, -1.314289, 1.570796, 1.552257],accel_mss,speed_ms,0,blend_radius_m)
  movel([-0.018169, -0.598052, -2.803126, -1.311210, 1.570796, 1.552627],accel_mss,speed_ms,0,blend_radius_m)
  movel([-0.017094, -0.600819, -2.802895, -1.308675, 1.570796, 1.553703],accel_mss,speed_ms,0,blend_radius_m)
  movel([-0.015272, -0.602944, -2.802715, -1.306731, 1.570796, 1.555524],accel_mss,speed_ms,0,blend_radius_m)
  movel([-0.012651, -0.604363, -2.802594, -1.305433, 1.570796, 1.558145],accel_mss,speed_ms,0,blend_radius_m)
  speed_ms = 0.005
  movel([-0.012651, -0.599373, -2.795777, -1.317239, 1.570796, 1.558145],accel_mss,speed_ms,0,blend_radius_m)
  speed_ms = 0.040
  movel([0.007037, -0.575986, -2.797664, -1.338739, 1.570796, 1.577833],accel_mss,speed_ms,0,blend_radius_m)
  speed_ms = 0.005
  movel([0.007037, -0.580592, -2.804518, -1.327280, 1.570796, 1.577833],accel_mss,speed_ms,0,blend_radius_m)
  speed_ms = 0.025
  movel([0.005993, -0.578452, -2.804680, -1.329257, 1.570796, 1.576790],accel_mss,speed_ms,0,blend_radius_m)
  movel([0.005278, -0.575976, -2.804865, -1.331548, 1.570796, 1.576075],accel_mss,speed_ms,0,blend_radius_m)
  movel([0.004895, -0.573193, -2.805071, -1.334125, 1.570796, 1.575691],accel_mss,speed_ms,0,blend_radius_m)
  movel([0.004846, -0.570117, -2.805294, -1.336977, 1.570796, 1.575642],accel_mss,speed_ms,0,blend_radius_m)
  movel([0.005129, -0.566780, -2.805533, -1.340076, 1.570796, 1.575925],accel_mss,speed_ms,0,blend_radius_m)
  movel([0.005755, -0.563194, -2.805784, -1.343411, 1.570796, 1.576551],accel_mss,speed_ms,0,blend_radius_m)
  movel([0.006728, -0.559376, -2.806047, -1.346967, 1.570796, 1.577525],accel_mss,speed_ms,0,blend_radius_m)
  movel([0.008047, -0.555360, -2.806316, -1.350713, 1.570796, 1.578844],accel_mss,speed_ms,0,blend_radius_m)
  movel([0.009716, -0.551162, -2.806592, -1.354636, 1.570796, 1.580513],accel_mss,speed_ms,0,blend_radius_m)
  movel([0.011747, -0.546797, -2.806871, -1.358721, 1.570796, 1.582543],accel_mss,speed_ms,0,blend_radius_m)
  movel([0.014131, -0.542307, -2.807150, -1.362931, 1.570796, 1.584927],accel_mss,speed_ms,0,blend_radius_m)
  movel([0.016885, -0.537695, -2.807430, -1.367264, 1.570796, 1.587681],accel_mss,speed_ms,0,blend_radius_m)
  movel([0.020006, -0.532992, -2.807706, -1.371691, 1.570796, 1.590802],accel_mss,speed_ms,0,blend_radius_m)
  movel([0.023499, -0.528224, -2.807978, -1.376187, 1.570796, 1.594295],accel_mss,speed_ms,0,blend_radius_m)
  movel([0.027365, -0.523419, -2.808243, -1.380727, 1.570796, 1.598161],accel_mss,speed_ms,0,blend_radius_m)
  movel([0.031600, -0.518605, -2.808500, -1.385284, 1.570796, 1.602396],accel_mss,speed_ms,0,blend_radius_m)
  movel([0.035938, -0.514103, -2.808733, -1.389553, 1.570796, 1.606734],accel_mss,speed_ms,0,blend_radius_m)
  movel([0.040340, -0.509939, -2.808941, -1.393509, 1.570796, 1.611137],accel_mss,speed_ms,0,blend_radius_m)
  movel([0.044769, -0.506121, -2.809127, -1.397142, 1.570796, 1.615565],accel_mss,speed_ms,0,blend_radius_m)
  movel([0.049204, -0.502652, -2.809291, -1.400447, 1.570796, 1.620000],accel_mss,speed_ms,0,blend_radius_m)
  movel([0.053607, -0.499540, -2.809434, -1.403415, 1.570796, 1.624403],accel_mss,speed_ms,0,blend_radius_m)
  movel([0.057938, -0.496805, -2.809557, -1.406027, 1.570796, 1.628734],accel_mss,speed_ms,0,blend_radius_m)
  movel([0.062180, -0.494431, -2.809661, -1.408297, 1.570796, 1.632976],accel_mss,speed_ms,0,blend_radius_m)
  movel([0.066279, -0.492447, -2.809747, -1.410195, 1.570796, 1.637075],accel_mss,speed_ms,0,blend_radius_m)
  movel([0.070217, -0.490847, -2.809815, -1.411727, 1.570796, 1.641013],accel_mss,speed_ms,0,blend_radius_m)
  movel([0.077485, -0.488806, -2.809901, -1.413683, 1.570796, 1.648281],accel_mss,speed_ms,0,blend_radius_m)
  movel([0.080741, -0.488382, -2.809918, -1.414089, 1.570796, 1.651537],accel_mss,speed_ms,0,blend_radius_m)
  movel([0.086385, -0.488705, -2.809905, -1.413779, 1.570796, 1.657181],accel_mss,speed_ms,0,blend_radius_m)
  movel([0.088712, -0.489452, -2.809874, -1.413063, 1.570796, 1.659508],accel_mss,speed_ms,0,blend_radius_m)
  movel([0.090669, -0.490594, -2.809826, -1.411970, 1.570796, 1.661466],accel_mss,speed_ms,0,blend_radius_m)
  speed_ms = 0.005
  movel([0.090669, -0.487553, -2.802869, -1.421967, 1.570796, 1.661466],accel_mss,speed_ms,0,blend_radius_m)
  speed_ms = 0.040
  movel([0.110623, -0.494154, -2.802583, -1.415652, 1.570796, 1.681419],accel_mss,speed_ms,0,blend_radius_m)
  speed_ms = 0.005
  movel([0.110623, -0.497318, -2.809534, -1.405537, 1.570796, 1.681419],accel_mss,speed_ms,0,blend_radius_m)
  speed_ms = 0.025
  movel([0.107860, -0.495328, -2.809622, -1.407439, 1.570796, 1.678657],accel_mss,speed_ms,0,blend_radius_m)
  movel([0.104297, -0.494386, -2.809663, -1.408340, 1.570796, 1.675093],accel_mss,speed_ms,0,blend_radius_m)
  movel([0.100017, -0.494472, -2.809659, -1.408257, 1.570796, 1.670814],accel_mss,speed_ms,0,blend_radius_m)
  movel([0.095095, -0.495569, -2.809611, -1.407209, 1.570796, 1.665891],accel_mss,speed_ms,0,blend_radius_m)
  movel([0.089640, -0.497634, -2.809520, -1.405236, 1.570796, 1.660436],accel_mss,speed_ms,0,blend_radius_m)
  movel([0.083731, -0.500645, -2.809383, -1.402361, 1.570796, 1.654527],accel_mss,speed_ms,0,blend_radius_m)
  movel([0.077480, -0.504557, -2.809201, -1.398631, 1.570796, 1.648276],accel_mss,speed_ms,0,blend_radius_m)
  movel([0.070971, -0.509334, -2.808971, -1.394084, 1.570796, 1.641768],accel_mss,speed_ms,0,blend_radius_m)
  movel([0.064325, -0.514920, -2.808691, -1.388778, 1.570796, 1.635121],accel_mss,speed_ms,0,blend_radius_m)
  movel([0.057700, -0.521200, -2.808363, -1.382826, 1.570796, 1.628496],accel_mss,speed_ms,0,blend_radius_m)
  movel([0.051361, -0.527945, -2.807993, -1.376450, 1.570796, 1.622157],accel_mss,speed_ms,0,blend_radius_m)
  movel([0.045580, -0.534930, -2.807593, -1.369866, 1.570796, 1.616376],accel_mss,speed_ms,0,blend_radius_m)
  movel([0.040590, -0.541955, -2.807172, -1.363262, 1.570796, 1.611386],accel_mss,speed_ms,0,blend_radius_m)
  movel([0.038474, -0.545412, -2.806958, -1.360019, 1.570796, 1.609271],accel_mss,speed_ms,0,blend_radius_m)
  movel([0.036641, -0.548801, -2.806744, -1.356844, 1.570796, 1.607438],accel_mss,speed_ms,0,blend_radius_m)
  movel([0.035120, -0.552103, -2.806531, -1.353756, 1.570796, 1.605917],accel_mss,speed_ms,0,blend_radius_m)
  movel([0.033946, -0.555293, -2.806321, -1.350776, 1.570796, 1.604742],accel_mss,speed_ms,0,blend_radius_m)
  movel([0.033135, -0.558347, -2.806116, -1.347926, 1.570796, 1.603931],accel_mss,speed_ms,0,blend_radius_m)
  movel([0.032727, -0.561233, -2.805920, -1.345236, 1.570796, 1.603523],accel_mss,speed_ms,0,blend_radius_m)
  speed_ms = 0.005
  movel([0.032727, -0.556950, -2.799039, -1.356399, 1.570796, 1.603523],accel_mss,speed_ms,0,blend_radius_m)
  speed_ms = 0.040
  movel([0.068280, -0.542322, -2.800000, -1.370067, 1.570796, 1.639077],accel_mss,speed_ms,0,blend_radius_m)
  speed_ms = 0.005
  movel([0.068280, -0.546352, -2.806899, -1.359138, 1.570796, 1.639077],accel_mss,speed_ms,0,blend_radius_m)
  speed_ms = 0.025
  movel([0.072553, -0.541253, -2.807215, -1.363921, 1.570796, 1.643349],accel_mss,speed_ms,0,blend_radius_m)
  movel([0.077095, -0.536482, -2.807502, -1.368406, 1.570796, 1.647891],accel_mss,speed_ms,0,blend_radius_m)
  movel([0.081825, -0.532070, -2.807759, -1.372559, 1.570796, 1.652622],accel_mss,speed_ms,0,blend_radius_m)
  movel([0.086644, -0.528075, -2.807986, -1.376328, 1.570796, 1.657440],accel_mss,speed_ms,0,blend_radius_m)
  movel([0.091459, -0.524534, -2.808182, -1.379673, 1.570796, 1.662255],accel_mss,speed_ms,0,blend_radius_m)
  movel([0.096168, -0.521491, -2.808347, -1.382551, 1.570796, 1.666964],accel_mss,speed_ms,0,blend_radius_m)
  movel([0.100686, -0.518985, -2.808480, -1.384924, 1.570796, 1.671482],accel_mss,speed_ms,0,blend_radius_m)
  movel([0.104903, -0.517061, -2.808581, -1.386747, 1.570796, 1.675699],accel_mss,speed_ms,0,blend_radius_m)
  movel([0.109483, -0.515668, -2.808653, -1.388068, 1.570796, 1.680280],accel_mss,speed_ms,0,blend_radius_m)
  movel([0.112978, -0.515528, -2.808660, -1.388201, 1.570796, 1.683775],accel_mss,speed_ms,0,blend_radius_m)
  movel([0.115503, -0.516508, -2.808609, -1.387272, 1.570796, 1.686299],accel_mss,speed_ms,0,blend_radius_m)
  movel([0.117149, -0.518488, -2.808506, -1.385395, 1.570796, 1.687946],accel_mss,speed_ms,0,blend_radius_m)
  movel([0.118032, -0.521321, -2.808356, -1.382711, 1.570796, 1.688829],accel_mss,speed_ms,0,blend_radius_m)
  movel([0.118264, -0.524884, -2.808163, -1.379342, 1.570796, 1.689060],accel_mss,speed_ms,0,blend_radius_m)
  movel([0.117953, -0.529039, -2.807932, -1.375418, 1.570796, 1.688749],accel_mss,speed_ms,0,blend_radius_m)
  movel([0.117219, -0.533648, -2.807668, -1.371073, 1.570796, 1.688015],accel_mss,speed_ms,0,blend_radius_m)
  speed_ms = 0.005
  movel([0.117219, -0.529838, -2.800754, -1.381797, 1.570796, 1.688015],accel_mss,speed_ms,0,blend_radius_m)
  speed_ms = 0.040
  movel([0.084510, -0.551516, -2.799406, -1.361467, 1.570796, 1.655307],accel_mss,speed_ms,0,blend_radius_m)
  speed_ms = 0.005
  movel([0.084510, -0.555706, -2.806293, -1.350390, 1.570796, 1.655307],accel_mss,speed_ms,0,blend_radius_m)
  speed_ms = 0.025
  movel([0.088925, -0.553047, -2.806469, -1.352873, 1.570796, 1.659721],accel_mss,speed_ms,0,blend_radius_m)
  movel([0.093004, -0.551013, -2.806601, -1.354774, 1.570796, 1.663801],accel_mss,speed_ms,0,blend_radius_m)
  movel([0.096743, -0.549595, -2.806693, -1.356101, 1.570796, 1.667540],accel_mss,speed_ms,0,blend_radius_m)
  movel([0.100140, -0.548753, -2.806747, -1.356889, 1.570796, 1.670936],accel_mss,speed_ms,0,blend_radius_m)
  movel([0.103191, -0.548467, -2.806765, -1.357157, 1.570796, 1.673988],accel_mss,speed_ms,0,blend_radius_m)
  movel([0.105893, -0.548706, -2.806750, -1.356933, 1.570796, 1.676690],accel_mss,speed_ms,0,blend_radius_m)
  movel([0.108253, -0.549436, -2.806703, -1.356250, 1.570796, 1.679049],accel_mss,speed_ms,0,blend_radius_m)
  movel([0.110260, -0.550640, -2.806625, -1.355124, 1.570796, 1.681057],accel_mss,speed_ms,0,blend_radius_m)
  movel([0.111933, -0.552272, -2.806520, -1.353598, 1.570796, 1.682729],accel_mss,speed_ms,0,blend_radius_m)
  movel([0.113269, -0.554301, -2.806386, -1.351701, 1.570796, 1.684066],accel_mss,speed_ms,0,blend_radius_m)
  movel([0.114270, -0.556703, -2.806227, -1.349460, 1.570796, 1.685066],accel_mss,speed_ms,0,blend_radius_m)
  movel([0.114947, -0.559434, -2.806043, -1.346913, 1.570796, 1.685743],accel_mss,speed_ms,0,blend_radius_m)
  movel([0.115302, -0.562468, -2.805835, -1.344086, 1.570796, 1.686098],accel_mss,speed_ms,0,blend_radius_m)
  movel([0.115078, -0.569299, -2.805353, -1.337736, 1.570796, 1.685874],accel_mss,speed_ms,0,blend_radius_m)
  movel([0.114508, -0.573038, -2.805082, -1.334269, 1.570796, 1.685305],accel_mss,speed_ms,0,blend_radius_m)
  movel([0.114176, -0.572179, -2.805145, -1.335065, 1.570796, 1.684972],accel_mss,speed_ms,0,blend_radius_m)
  speed_ms = 0.005
  movel([0.114176, -0.567712, -2.798280, -1.346397, 1.570796, 1.684972],accel_mss,speed_ms,0,blend_radius_m)
  speed_ms = 0.040
  movel([0.141519, -0.562009, -2.798688, -1.351692, 1.570796, 1.712316],accel_mss,speed_ms,0,blend_radius_m)
  speed_ms = 0.005
  movel([0.141519, -0.566379, -2.805561, -1.340449, 1.570796, 1.712316],accel_mss,speed_ms,0,blend_radius_m)
  speed_ms = 0.025
  movel([0.137715, -0.572995, -2.805085, -1.334308, 1.570796, 1.708512],accel_mss,speed_ms,0,blend_radius_m)
  movel([0.134491, -0.579437, -2.804605, -1.328347, 1.570796, 1.705287],accel_mss,speed_ms,0,blend_radius_m)
  movel([0.131717, -0.585709, -2.804122, -1.322557, 1.570796, 1.702514],accel_mss,speed_ms,0,blend_radius_m)
  movel([0.129255, -0.591825, -2.803637, -1.316927, 1.570796, 1.700051],accel_mss,speed_ms,0,blend_radius_m)
  movel([0.126862, -0.598387, -2.803099, -1.310903, 1.570796, 1.697659],accel_mss,speed_ms,0,blend_radius_m)
  movel([0.125961, -0.601487, -2.802838, -1.308063, 1.570796, 1.696757],accel_mss,speed_ms,0,blend_radius_m)
  movel([0.125376, -0.604382, -2.802592, -1.305415, 1.570796, 1.696173],accel_mss,speed_ms,0,blend_radius_m)
  movel([0.125184, -0.607002, -2.802366, -1.303021, 1.570796, 1.695980],accel_mss,speed_ms,0,blend_radius_m)
  movel([0.125467, -0.609223, -2.802172, -1.300993, 1.570796, 1.696263],accel_mss,speed_ms,0,blend_radius_m)
  movel([0.126291, -0.610890, -2.802026, -1.299474, 1.570796, 1.697088],accel_mss,speed_ms,0,blend_radius_m)
  movel([0.127710, -0.611876, -2.801938, -1.298575, 1.570796, 1.698506],accel_mss,speed_ms,0,blend_radius_m)
  movel([0.130856, -0.612205, -2.801909, -1.298275, 1.570796, 1.701652],accel_mss,speed_ms,0,blend_radius_m)
  movel([0.132407, -0.612389, -2.801893, -1.298108, 1.570796, 1.703203],accel_mss,speed_ms,0,blend_radius_m)
  movel([0.133647, -0.612982, -2.801840, -1.297567, 1.570796, 1.704444],accel_mss,speed_ms,0,blend_radius_m)
  movel([0.134411, -0.614473, -2.801706, -1.296210, 1.570796, 1.705207],accel_mss,speed_ms,0,blend_radius_m)
  movel([0.134534, -0.616777, -2.801499, -1.294114, 1.570796, 1.705330],accel_mss,speed_ms,0,blend_radius_m)
  movel([0.134155, -0.619680, -2.801233, -1.291475, 1.570796, 1.704951],accel_mss,speed_ms,0,blend_radius_m)
  movel([0.133404, -0.622971, -2.800928, -1.288489, 1.570796, 1.704200],accel_mss,speed_ms,0,blend_radius_m)
  movel([0.131302, -0.629899, -2.800272, -1.282218, 1.570796, 1.702098],accel_mss,speed_ms,0,blend_radius_m)
  movel([0.124391, -0.649574, -2.798299, -1.264516, 1.570796, 1.695188],accel_mss,speed_ms,0,blend_radius_m)
  movel([0.119712, -0.663005, -2.796857, -1.252527, 1.570796, 1.690508],accel_mss,speed_ms,0,blend_radius_m)
  movel([0.118564, -0.666973, -2.796416, -1.249000, 1.570796, 1.689361],accel_mss,speed_ms,0,blend_radius_m)
  movel([0.117618, -0.671063, -2.795954, -1.245372, 1.570796, 1.688415],accel_mss,speed_ms,0,blend_radius_m)
  movel([0.116433, -0.679241, -2.795009, -1.238138, 1.570796, 1.687230],accel_mss,speed_ms,0,blend_radius_m)
  movel([0.116251, -0.683150, -2.794547, -1.234692, 1.570796, 1.687047],accel_mss,speed_ms,0,blend_radius_m)
  movel([0.116378, -0.686816, -2.794108, -1.231466, 1.570796, 1.687175],accel_mss,speed_ms,0,blend_radius_m)
  movel([0.116838, -0.690154, -2.793702, -1.228533, 1.570796, 1.687635],accel_mss,speed_ms,0,blend_radius_m)
  movel([0.117658, -0.693082, -2.793342, -1.225965, 1.570796, 1.688454],accel_mss,speed_ms,0,blend_radius_m)
  movel([0.118866, -0.695499, -2.793042, -1.223848, 1.570796, 1.689662],accel_mss,speed_ms,0,blend_radius_m)
  movel([0.120484, -0.697338, -2.792812, -1.222239, 1.570796, 1.691280],accel_mss,speed_ms,0,blend_radius_m)
  movel([0.122549, -0.698494, -2.792667, -1.221228, 1.570796, 1.693346],accel_mss,speed_ms,0,blend_radius_m)
  movel([0.125089, -0.698888, -2.792617, -1.220884, 1.570796, 1.695885],accel_mss,speed_ms,0,blend_radius_m)
  movel([0.128131, -0.698428, -2.792675, -1.221286, 1.570796, 1.698928],accel_mss,speed_ms,0,blend_radius_m)
  movel([0.131721, -0.697017, -2.792852, -1.222519, 1.570796, 1.702517],accel_mss,speed_ms,0,blend_radius_m)
  movel([0.135894, -0.694563, -2.793159, -1.224667, 1.570796, 1.706690],accel_mss,speed_ms,0,blend_radius_m)
  movel([0.140697, -0.690962, -2.793603, -1.227824, 1.570796, 1.711493],accel_mss,speed_ms,0,blend_radius_m)
  movel([0.144464, -0.687665, -2.794005, -1.230719, 1.570796, 1.715261],accel_mss,speed_ms,0,blend_radius_m)
  movel([0.148149, -0.684073, -2.794437, -1.233879, 1.570796, 1.718945],accel_mss,speed_ms,0,blend_radius_m)
  movel([0.151771, -0.680225, -2.794894, -1.237270, 1.570796, 1.722567],accel_mss,speed_ms,0,blend_radius_m)
  movel([0.155340, -0.676172, -2.795367, -1.240850, 1.570796, 1.726136],accel_mss,speed_ms,0,blend_radius_m)
  movel([0.162365, -0.667650, -2.796340, -1.248399, 1.570796, 1.733161],accel_mss,speed_ms,0,blend_radius_m)
  movel([0.169324, -0.658907, -2.797305, -1.256177, 1.570796, 1.740120],accel_mss,speed_ms,0,blend_radius_m)
  movel([0.176535, -0.650139, -2.798240, -1.264011, 1.570796, 1.747331],accel_mss,speed_ms,0,blend_radius_m)
  movel([0.180311, -0.645826, -2.798687, -1.267876, 1.570796, 1.751107],accel_mss,speed_ms,0,blend_radius_m)
  movel([0.184177, -0.641674, -2.799111, -1.271604, 1.570796, 1.754973],accel_mss,speed_ms,0,blend_radius_m)
  movel([0.188111, -0.637756, -2.799504, -1.275130, 1.570796, 1.758907],accel_mss,speed_ms,0,blend_radius_m)
  movel([0.192093, -0.634163, -2.799858, -1.278368, 1.570796, 1.762889],accel_mss,speed_ms,0,blend_radius_m)
  movel([0.196091, -0.630981, -2.800168, -1.281240, 1.570796, 1.766888],accel_mss,speed_ms,0,blend_radius_m)
  movel([0.200089, -0.628297, -2.800426, -1.283667, 1.570796, 1.770885],accel_mss,speed_ms,0,blend_radius_m)
  movel([0.208531, -0.623802, -2.800851, -1.287736, 1.570796, 1.779327],accel_mss,speed_ms,0,blend_radius_m)
  movel([0.211406, -0.622083, -2.801011, -1.289295, 1.570796, 1.782202],accel_mss,speed_ms,0,blend_radius_m)
  movel([0.214435, -0.619847, -2.801218, -1.291324, 1.570796, 1.785231],accel_mss,speed_ms,0,blend_radius_m)
  movel([0.217463, -0.617079, -2.801471, -1.293839, 1.570796, 1.788260],accel_mss,speed_ms,0,blend_radius_m)
  movel([0.220197, -0.613942, -2.801754, -1.296693, 1.570796, 1.790993],accel_mss,speed_ms,0,blend_radius_m)
  movel([0.221366, -0.612277, -2.801903, -1.298209, 1.570796, 1.792163],accel_mss,speed_ms,0,blend_radius_m)
  movel([0.222353, -0.610578, -2.802053, -1.299758, 1.570796, 1.793150],accel_mss,speed_ms,0,blend_radius_m)
  speed_ms = 0.005
  movel([0.222353, -0.605491, -2.795247, -1.311652, 1.570796, 1.793150],accel_mss,speed_ms,0,blend_radius_m)
  speed_ms = 0.040
  movel([0.236641, -0.575239, -2.797721, -1.339429, 1.570796, 1.807437],accel_mss,speed_ms,0,blend_radius_m)
  speed_ms = 0.005
  movel([0.236641, -0.579832, -2.804575, -1.327982, 1.570796, 1.807437],accel_mss,speed_ms,0,blend_radius_m)
  speed_ms = 0.025
  movel([0.237599, -0.579729, -2.804583, -1.328076, 1.570796, 1.808395],accel_mss,speed_ms,0,blend_radius_m)
  movel([0.237681, -0.580741, -2.804506, -1.327142, 1.570796, 1.808477],accel_mss,speed_ms,0,blend_radius_m)
  movel([0.237034, -0.582361, -2.804382, -1.325646, 1.570796, 1.807830],accel_mss,speed_ms,0,blend_radius_m)
  movel([0.235833, -0.584077, -2.804250, -1.324063, 1.570796, 1.806629],accel_mss,speed_ms,0,blend_radius_m)
  movel([0.234372, -0.585507, -2.804138, -1.322744, 1.570796, 1.805169],accel_mss,speed_ms,0,blend_radius_m)
  movel([0.232871, -0.586684, -2.804046, -1.321659, 1.570796, 1.803667],accel_mss,speed_ms,0,blend_radius_m)
  movel([0.229848, -0.588769, -2.803881, -1.319739, 1.570796, 1.800644],accel_mss,speed_ms,0,blend_radius_m)
  movel([0.227666, -0.590488, -2.803744, -1.318157, 1.570796, 1.798462],accel_mss,speed_ms,0,blend_radius_m)
  movel([0.225527, -0.592444, -2.803587, -1.316359, 1.570796, 1.796324],accel_mss,speed_ms,0,blend_radius_m)
  movel([0.221382, -0.596891, -2.803223, -1.312275, 1.570796, 1.792179],accel_mss,speed_ms,0,blend_radius_m)
  movel([0.217443, -0.601772, -2.802814, -1.307803, 1.570796, 1.788239],accel_mss,speed_ms,0,blend_radius_m)
  movel([0.213738, -0.606728, -2.802390, -1.303271, 1.570796, 1.784534],accel_mss,speed_ms,0,blend_radius_m)
  movel([0.212904, -0.607944, -2.802284, -1.302161, 1.570796, 1.783700],accel_mss,speed_ms,0,blend_radius_m)
  movel([0.212415, -0.609046, -2.802188, -1.301155, 1.570796, 1.783211],accel_mss,speed_ms,0,blend_radius_m)
  movel([0.212668, -0.609742, -2.802127, -1.300521, 1.570796, 1.783465],accel_mss,speed_ms,0,blend_radius_m)
  movel([0.213509, -0.609803, -2.802121, -1.300464, 1.570796, 1.784306],accel_mss,speed_ms,0,blend_radius_m)
  movel([0.215716, -0.609347, -2.802162, -1.300881, 1.570796, 1.786513],accel_mss,speed_ms,0,blend_radius_m)
  movel([0.218137, -0.608446, -2.802240, -1.301703, 1.570796, 1.788934],accel_mss,speed_ms,0,blend_radius_m)
  movel([0.220731, -0.607137, -2.802354, -1.302898, 1.570796, 1.791528],accel_mss,speed_ms,0,blend_radius_m)
  movel([0.223452, -0.605439, -2.802501, -1.304448, 1.570796, 1.794249],accel_mss,speed_ms,0,blend_radius_m)
  movel([0.226242, -0.603405, -2.802676, -1.306308, 1.570796, 1.797038],accel_mss,speed_ms,0,blend_radius_m)
  movel([0.229059, -0.601049, -2.802875, -1.308464, 1.570796, 1.799856],accel_mss,speed_ms,0,blend_radius_m)
  movel([0.231847, -0.598417, -2.803096, -1.310876, 1.570796, 1.802643],accel_mss,speed_ms,0,blend_radius_m)
  movel([0.234561, -0.595529, -2.803335, -1.313525, 1.570796, 1.805357],accel_mss,speed_ms,0,blend_radius_m)
  movel([0.234154, -0.597105, -2.803205, -1.312079, 1.570796, 1.804950],accel_mss,speed_ms,0,blend_radius_m)
  movel([0.234464, -0.598118, -2.803121, -1.311150, 1.570796, 1.805260],accel_mss,speed_ms,0,blend_radius_m)
  movel([0.235344, -0.598533, -2.803086, -1.310770, 1.570796, 1.806141],accel_mss,speed_ms,0,blend_radius_m)
  movel([0.236639, -0.598317, -2.803104, -1.310967, 1.570796, 1.807436],accel_mss,speed_ms,0,blend_radius_m)
  movel([0.238175, -0.597544, -2.803169, -1.311676, 1.570796, 1.808971],accel_mss,speed_ms,0,blend_radius_m)
  movel([0.239829, -0.596394, -2.803264, -1.312731, 1.570796, 1.810626],accel_mss,speed_ms,0,blend_radius_m)
  movel([0.243225, -0.593414, -2.803508, -1.315467, 1.570796, 1.814021],accel_mss,speed_ms,0,blend_radius_m)
  movel([0.247467, -0.589044, -2.803859, -1.319486, 1.570796, 1.818263],accel_mss,speed_ms,0,blend_radius_m)
  movel([0.251492, -0.584297, -2.804233, -1.323859, 1.570796, 1.822288],accel_mss,speed_ms,0,blend_radius_m)
  movel([0.255190, -0.579317, -2.804614, -1.328457, 1.570796, 1.825986],accel_mss,speed_ms,0,blend_radius_m)
  movel([0.258444, -0.574244, -2.804994, -1.333152, 1.570796, 1.829240],accel_mss,speed_ms,0,blend_radius_m)
  movel([0.259355, -0.572554, -2.805118, -1.334717, 1.570796, 1.830151],accel_mss,speed_ms,0,blend_radius_m)
  movel([0.259738, -0.571157, -2.805219, -1.336012, 1.570796, 1.830534],accel_mss,speed_ms,0,blend_radius_m)
  movel([0.259411, -0.570523, -2.805265, -1.336601, 1.570796, 1.830208],accel_mss,speed_ms,0,blend_radius_m)
  movel([0.258704, -0.570314, -2.805280, -1.336794, 1.570796, 1.829501],accel_mss,speed_ms,0,blend_radius_m)
  movel([0.255838, -0.570359, -2.805277, -1.336753, 1.570796, 1.826635],accel_mss,speed_ms,0,blend_radius_m)
  movel([0.250064, -0.571195, -2.805216, -1.335977, 1.570796, 1.820861],accel_mss,speed_ms,0,blend_radius_m)
  movel([0.247550, -0.570705, -2.805252, -1.336432, 1.570796, 1.818347],accel_mss,speed_ms,0,blend_radius_m)
  movel([0.252228, -0.564899, -2.805665, -1.341824, 1.570796, 1.823024],accel_mss,speed_ms,0,blend_radius_m)
  movel([0.254770, -0.562220, -2.805852, -1.344317, 1.570796, 1.825566],accel_mss,speed_ms,0,blend_radius_m)
  movel([0.257396, -0.559847, -2.806015, -1.346528, 1.570796, 1.828193],accel_mss,speed_ms,0,blend_radius_m)
  movel([0.259201, -0.558496, -2.806106, -1.347787, 1.570796, 1.829998],accel_mss,speed_ms,0,blend_radius_m)
  movel([0.261070, -0.557330, -2.806185, -1.348874, 1.570796, 1.831866],accel_mss,speed_ms,0,blend_radius_m)
  movel([0.264381, -0.555873, -2.806282, -1.350233, 1.570796, 1.835178],accel_mss,speed_ms,0,blend_radius_m)
  movel([0.266059, -0.555934, -2.806278, -1.350177, 1.570796, 1.836855],accel_mss,speed_ms,0,blend_radius_m)
  movel([0.266502, -0.556460, -2.806243, -1.349686, 1.570796, 1.837298],accel_mss,speed_ms,0,blend_radius_m)
  movel([0.266569, -0.557356, -2.806183, -1.348850, 1.570796, 1.837365],accel_mss,speed_ms,0,blend_radius_m)
  movel([0.266060, -0.558947, -2.806076, -1.347367, 1.570796, 1.836856],accel_mss,speed_ms,0,blend_radius_m)
  movel([0.265041, -0.560765, -2.805952, -1.345672, 1.570796, 1.835837],accel_mss,speed_ms,0,blend_radius_m)
  movel([0.262212, -0.564544, -2.805690, -1.342154, 1.570796, 1.833008],accel_mss,speed_ms,0,blend_radius_m)
  speed_ms = 0.005
  movel([0.262212, -0.560206, -2.798814, -1.353369, 1.570796, 1.833008],accel_mss,speed_ms,0,blend_radius_m)
  speed_ms = 0.040
  movel([0.290577, -0.451763, -2.804141, -1.456485, 1.570796, 1.861374],accel_mss,speed_ms,0,blend_radius_m)
  speed_ms = 0.005
  movel([0.290577, -0.454128, -2.811123, -1.447138, 1.570796, 1.861374],accel_mss,speed_ms,0,blend_radius_m)
  speed_ms = 0.025
  movel([0.292801, -0.451970, -2.811185, -1.449234, 1.570796, 1.863598],accel_mss,speed_ms,0,blend_radius_m)
  movel([0.295031, -0.450106, -2.811237, -1.451045, 1.570796, 1.865827],accel_mss,speed_ms,0,blend_radius_m)
  movel([0.297215, -0.448552, -2.811280, -1.452557, 1.570796, 1.868012],accel_mss,speed_ms,0,blend_radius_m)
  movel([0.301288, -0.446409, -2.811337, -1.454643, 1.570796, 1.872084],accel_mss,speed_ms,0,blend_radius_m)
  movel([0.303082, -0.445841, -2.811352, -1.455196, 1.570796, 1.873879],accel_mss,speed_ms,0,blend_radius_m)
  movel([0.305963, -0.445766, -2.811354, -1.455269, 1.570796, 1.876760],accel_mss,speed_ms,0,blend_radius_m)
  movel([0.307802, -0.446975, -2.811322, -1.454091, 1.570796, 1.878598],accel_mss,speed_ms,0,blend_radius_m)
  movel([0.308768, -0.449144, -2.811264, -1.451982, 1.570796, 1.879564],accel_mss,speed_ms,0,blend_radius_m)
  movel([0.309023, -0.452029, -2.811184, -1.449176, 1.570796, 1.879819],accel_mss,speed_ms,0,blend_radius_m)
  movel([0.308729, -0.455391, -2.811086, -1.445911, 1.570796, 1.879525],accel_mss,speed_ms,0,blend_radius_m)
  movel([0.307527, -0.461057, -2.810914, -1.440418, 1.570796, 1.878323],accel_mss,speed_ms,0,blend_radius_m)
  movel([0.305534, -0.467274, -2.810711, -1.434404, 1.570796, 1.876330],accel_mss,speed_ms,0,blend_radius_m)
  movel([0.302802, -0.473924, -2.810478, -1.427986, 1.570796, 1.873598],accel_mss,speed_ms,0,blend_radius_m)
  movel([0.296051, -0.487526, -2.809953, -1.414910, 1.570796, 1.866847],accel_mss,speed_ms,0,blend_radius_m)
  movel([0.295041, -0.490393, -2.809834, -1.412162, 1.570796, 1.865837],accel_mss,speed_ms,0,blend_radius_m)
  movel([0.294976, -0.492539, -2.809743, -1.410107, 1.570796, 1.865773],accel_mss,speed_ms,0,blend_radius_m)
  movel([0.295867, -0.493557, -2.809699, -1.409133, 1.570796, 1.866664],accel_mss,speed_ms,0,blend_radius_m)
  movel([0.297298, -0.493961, -2.809682, -1.408746, 1.570796, 1.868094],accel_mss,speed_ms,0,blend_radius_m)
  movel([0.298841, -0.494248, -2.809669, -1.408472, 1.570796, 1.869638],accel_mss,speed_ms,0,blend_radius_m)
  movel([0.300053, -0.494926, -2.809640, -1.407824, 1.570796, 1.870850],accel_mss,speed_ms,0,blend_radius_m)
  movel([0.300567, -0.496154, -2.809586, -1.406649, 1.570796, 1.871363],accel_mss,speed_ms,0,blend_radius_m)
  movel([0.300568, -0.497871, -2.809509, -1.405009, 1.570796, 1.871364],accel_mss,speed_ms,0,blend_radius_m)
  movel([0.299667, -0.502072, -2.809317, -1.401000, 1.570796, 1.870463],accel_mss,speed_ms,0,blend_radius_m)
  movel([0.297719, -0.508533, -2.809010, -1.394846, 1.570796, 1.868515],accel_mss,speed_ms,0,blend_radius_m)
  movel([0.295397, -0.515209, -2.808676, -1.388504, 1.570796, 1.866193],accel_mss,speed_ms,0,blend_radius_m)
  movel([0.292707, -0.522068, -2.808316, -1.382005, 1.570796, 1.863504],accel_mss,speed_ms,0,blend_radius_m)
  movel([0.289682, -0.529078, -2.807930, -1.375381, 1.570796, 1.860478],accel_mss,speed_ms,0,blend_radius_m)
  movel([0.286334, -0.536200, -2.807518, -1.368671, 1.570796, 1.857130],accel_mss,speed_ms,0,blend_radius_m)
  movel([0.282693, -0.543398, -2.807083, -1.361908, 1.570796, 1.853490],accel_mss,speed_ms,0,blend_radius_m)
  movel([0.278762, -0.550651, -2.806625, -1.355113, 1.570796, 1.849559],accel_mss,speed_ms,0,blend_radius_m)
  movel([0.274569, -0.557927, -2.806145, -1.348317, 1.570796, 1.845366],accel_mss,speed_ms,0,blend_radius_m)
  movel([0.271720, -0.562531, -2.805830, -1.344028, 1.570796, 1.842516],accel_mss,speed_ms,0,blend_radius_m)
  movel([0.268543, -0.567103, -2.805510, -1.339776, 1.570796, 1.839339],accel_mss,speed_ms,0,blend_radius_m)
  movel([0.265062, -0.571326, -2.805207, -1.335856, 1.570796, 1.835858],accel_mss,speed_ms,0,blend_radius_m)
  movel([0.263216, -0.573199, -2.805070, -1.334120, 1.570796, 1.834012],accel_mss,speed_ms,0,blend_radius_m)
  movel([0.261298, -0.574873, -2.804947, -1.332569, 1.570796, 1.832094],accel_mss,speed_ms,0,blend_radius_m)
  speed_ms = 0.005
  movel([0.261298, -0.570362, -2.798086, -1.343941, 1.570796, 1.832094],accel_mss,speed_ms,0,blend_radius_m)
  speed_ms = 0.040
  movel([0.251459, -0.583325, -2.797096, -1.331968, 1.570796, 1.822256],accel_mss,speed_ms,0,blend_radius_m)
  speed_ms = 0.005
  movel([0.251459, -0.588052, -2.803938, -1.320399, 1.570796, 1.822256],accel_mss,speed_ms,0,blend_radius_m)
  speed_ms = 0.025
  movel([0.251817, -0.588872, -2.803873, -1.319644, 1.570796, 1.822613],accel_mss,speed_ms,0,blend_radius_m)
  movel([0.251535, -0.590251, -2.803763, -1.318375, 1.570796, 1.822332],accel_mss,speed_ms,0,blend_radius_m)
  movel([0.250759, -0.591940, -2.803627, -1.316822, 1.570796, 1.821556],accel_mss,speed_ms,0,blend_radius_m)
  movel([0.249620, -0.593689, -2.803485, -1.315214, 1.570796, 1.820416],accel_mss,speed_ms,0,blend_radius_m)
  movel([0.247973, -0.595546, -2.803334, -1.313510, 1.570796, 1.818769],accel_mss,speed_ms,0,blend_radius_m)
  movel([0.246257, -0.597087, -2.803207, -1.312095, 1.570796, 1.817054],accel_mss,speed_ms,0,blend_radius_m)
  movel([0.244576, -0.598544, -2.803086, -1.310759, 1.570796, 1.815372],accel_mss,speed_ms,0,blend_radius_m)
  movel([0.243054, -0.600140, -2.802952, -1.309297, 1.570796, 1.813850],accel_mss,speed_ms,0,blend_radius_m)
  movel([0.241521, -0.602666, -2.802739, -1.306985, 1.570796, 1.812318],accel_mss,speed_ms,0,blend_radius_m)
  movel([0.240827, -0.603963, -2.802628, -1.305798, 1.570796, 1.811624],accel_mss,speed_ms,0,blend_radius_m)
  movel([0.239860, -0.605377, -2.802507, -1.304505, 1.570796, 1.810656],accel_mss,speed_ms,0,blend_radius_m)
  movel([0.236774, -0.608999, -2.802192, -1.301198, 1.570796, 1.807570],accel_mss,speed_ms,0,blend_radius_m)
  movel([0.233629, -0.612196, -2.801910, -1.298283, 1.570796, 1.804425],accel_mss,speed_ms,0,blend_radius_m)
  movel([0.230406, -0.615035, -2.801656, -1.295698, 1.570796, 1.801202],accel_mss,speed_ms,0,blend_radius_m)
  movel([0.227084, -0.617610, -2.801423, -1.293356, 1.570796, 1.797880],accel_mss,speed_ms,0,blend_radius_m)
  movel([0.228805, -0.616122, -2.801558, -1.294710, 1.570796, 1.799602],accel_mss,speed_ms,0,blend_radius_m)
  movel([0.230513, -0.614870, -2.801671, -1.295848, 1.570796, 1.801309],accel_mss,speed_ms,0,blend_radius_m)
  movel([0.232068, -0.614186, -2.801732, -1.296471, 1.570796, 1.802864],accel_mss,speed_ms,0,blend_radius_m)
  movel([0.233072, -0.614438, -2.801710, -1.296242, 1.570796, 1.803869],accel_mss,speed_ms,0,blend_radius_m)
  movel([0.233129, -0.615709, -2.801595, -1.295084, 1.570796, 1.803926],accel_mss,speed_ms,0,blend_radius_m)
  movel([0.232407, -0.617510, -2.801432, -1.293447, 1.570796, 1.803204],accel_mss,speed_ms,0,blend_radius_m)
  movel([0.231176, -0.619417, -2.801257, -1.291715, 1.570796, 1.801972],accel_mss,speed_ms,0,blend_radius_m)
  movel([0.227244, -0.624119, -2.800821, -1.287449, 1.570796, 1.798040],accel_mss,speed_ms,0,blend_radius_m)
  movel([0.224667, -0.626784, -2.800570, -1.285035, 1.570796, 1.795463],accel_mss,speed_ms,0,blend_radius_m)
  movel([0.222039, -0.629222, -2.800337, -1.282830, 1.570796, 1.792836],accel_mss,speed_ms,0,blend_radius_m)
  movel([0.219385, -0.631405, -2.800127, -1.280857, 1.570796, 1.790182],accel_mss,speed_ms,0,blend_radius_m)
  movel([0.222400, -0.629296, -2.800330, -1.282763, 1.570796, 1.793197],accel_mss,speed_ms,0,blend_radius_m)
  movel([0.225548, -0.626766, -2.800571, -1.285052, 1.570796, 1.796345],accel_mss,speed_ms,0,blend_radius_m)
  movel([0.228636, -0.624343, -2.800800, -1.287246, 1.570796, 1.799433],accel_mss,speed_ms,0,blend_radius_m)
  movel([0.231471, -0.622537, -2.800969, -1.288883, 1.570796, 1.802267],accel_mss,speed_ms,0,blend_radius_m)
  movel([0.232257, -0.622347, -2.800987, -1.289055, 1.570796, 1.803053],accel_mss,speed_ms,0,blend_radius_m)
  movel([0.232280, -0.622863, -2.800939, -1.288587, 1.570796, 1.803076],accel_mss,speed_ms,0,blend_radius_m)
  movel([0.230688, -0.625909, -2.800653, -1.285828, 1.570796, 1.801484],accel_mss,speed_ms,0,blend_radius_m)
  movel([0.229209, -0.628173, -2.800438, -1.283779, 1.570796, 1.800006],accel_mss,speed_ms,0,blend_radius_m)
  movel([0.227550, -0.630385, -2.800225, -1.281779, 1.570796, 1.798346],accel_mss,speed_ms,0,blend_radius_m)
  movel([0.225753, -0.632485, -2.800022, -1.279882, 1.570796, 1.796549],accel_mss,speed_ms,0,blend_radius_m)
  movel([0.226667, -0.631634, -2.800105, -1.280651, 1.570796, 1.797464],accel_mss,speed_ms,0,blend_radius_m)
  movel([0.227692, -0.630934, -2.800172, -1.281283, 1.570796, 1.798488],accel_mss,speed_ms,0,blend_radius_m)
  movel([0.229931, -0.629969, -2.800265, -1.282155, 1.570796, 1.800727],accel_mss,speed_ms,0,blend_radius_m)
  movel([0.232159, -0.629581, -2.800303, -1.282505, 1.570796, 1.802955],accel_mss,speed_ms,0,blend_radius_m)
  movel([0.234085, -0.629746, -2.800287, -1.282356, 1.570796, 1.804882],accel_mss,speed_ms,0,blend_radius_m)
  movel([0.235424, -0.630434, -2.800221, -1.281734, 1.570796, 1.806220],accel_mss,speed_ms,0,blend_radius_m)
  movel([0.235885, -0.631608, -2.800107, -1.280673, 1.570796, 1.806681],accel_mss,speed_ms,0,blend_radius_m)
  movel([0.235698, -0.632368, -2.800033, -1.279988, 1.570796, 1.806495],accel_mss,speed_ms,0,blend_radius_m)
  movel([0.235185, -0.633232, -2.799949, -1.279207, 1.570796, 1.805982],accel_mss,speed_ms,0,blend_radius_m)
  movel([0.234317, -0.634206, -2.799854, -1.278329, 1.570796, 1.805113],accel_mss,speed_ms,0,blend_radius_m)
  movel([0.233049, -0.635280, -2.799749, -1.277361, 1.570796, 1.803845],accel_mss,speed_ms,0,blend_radius_m)
  movel([0.231643, -0.636132, -2.799665, -1.276592, 1.570796, 1.802439],accel_mss,speed_ms,0,blend_radius_m)
  movel([0.226386, -0.637686, -2.799511, -1.275193, 1.570796, 1.797183],accel_mss,speed_ms,0,blend_radius_m)
  movel([0.224340, -0.638400, -2.799439, -1.274549, 1.570796, 1.795136],accel_mss,speed_ms,0,blend_radius_m)
  movel([0.222146, -0.639530, -2.799326, -1.273533, 1.570796, 1.792942],accel_mss,speed_ms,0,blend_radius_m)
  movel([0.218320, -0.642349, -2.799042, -1.270998, 1.570796, 1.789117],accel_mss,speed_ms,0,blend_radius_m)
  movel([0.214469, -0.645422, -2.798729, -1.268239, 1.570796, 1.785265],accel_mss,speed_ms,0,blend_radius_m)
  movel([0.212548, -0.646675, -2.798600, -1.267114, 1.570796, 1.783344],accel_mss,speed_ms,0,blend_radius_m)
  movel([0.210756, -0.647498, -2.798515, -1.266376, 1.570796, 1.781552],accel_mss,speed_ms,0,blend_radius_m)
  movel([0.209315, -0.647694, -2.798494, -1.266200, 1.570796, 1.780111],accel_mss,speed_ms,0,blend_radius_m)
  movel([0.208440, -0.647079, -2.798558, -1.266752, 1.570796, 1.779236],accel_mss,speed_ms,0,blend_radius_m)
  movel([0.210303, -0.644467, -2.798827, -1.269095, 1.570796, 1.781100],accel_mss,speed_ms,0,blend_radius_m)
  movel([0.212339, -0.641934, -2.799084, -1.271371, 1.570796, 1.783136],accel_mss,speed_ms,0,blend_radius_m)
  speed_ms = 0.005
  movel([0.212339, -0.636366, -2.792334, -1.283689, 1.570796, 1.783136],accel_mss,speed_ms,0,blend_radius_m)
  speed_ms = 0.040
  movel([0.230373, -0.641563, -2.791804, -1.279022, 1.570796, 1.801169],accel_mss,speed_ms,0,blend_radius_m)
  speed_ms = 0.005
  movel([0.230373, -0.647209, -2.798545, -1.266636, 1.570796, 1.801169],accel_mss,speed_ms,0,blend_radius_m)
  speed_ms = 0.025
  movel([0.231696, -0.645339, -2.798737, -1.268313, 1.570796, 1.802492],accel_mss,speed_ms,0,blend_radius_m)
  movel([0.233355, -0.643804, -2.798894, -1.269691, 1.570796, 1.804152],accel_mss,speed_ms,0,blend_radius_m)
  movel([0.235068, -0.642757, -2.799001, -1.270631, 1.570796, 1.805864],accel_mss,speed_ms,0,blend_radius_m)
  movel([0.236535, -0.642364, -2.799041, -1.270984, 1.570796, 1.807332],accel_mss,speed_ms,0,blend_radius_m)
  movel([0.237599, -0.642606, -2.799016, -1.270767, 1.570796, 1.808396],accel_mss,speed_ms,0,blend_radius_m)
  movel([0.238355, -0.643262, -2.798950, -1.270177, 1.570796, 1.809151],accel_mss,speed_ms,0,blend_radius_m)
  movel([0.239319, -0.645238, -2.798748, -1.268403, 1.570796, 1.810115],accel_mss,speed_ms,0,blend_radius_m)
  movel([0.240486, -0.643023, -2.798974, -1.270392, 1.570796, 1.811283],accel_mss,speed_ms,0,blend_radius_m)
  movel([0.241179, -0.640966, -2.799182, -1.272241, 1.570796, 1.811976],accel_mss,speed_ms,0,blend_radius_m)
  movel([0.241343, -0.639243, -2.799355, -1.273791, 1.570796, 1.812139],accel_mss,speed_ms,0,blend_radius_m)
  movel([0.240949, -0.637998, -2.799479, -1.274911, 1.570796, 1.811745],accel_mss,speed_ms,0,blend_radius_m)
  movel([0.241923, -0.638204, -2.799459, -1.274726, 1.570796, 1.812719],accel_mss,speed_ms,0,blend_radius_m)
  movel([0.242636, -0.638737, -2.799406, -1.274246, 1.570796, 1.813433],accel_mss,speed_ms,0,blend_radius_m)
  movel([0.243413, -0.640569, -2.799222, -1.272598, 1.570796, 1.814209],accel_mss,speed_ms,0,blend_radius_m)
  movel([0.243579, -0.643072, -2.798969, -1.270348, 1.570796, 1.814375],accel_mss,speed_ms,0,blend_radius_m)
  movel([0.243396, -0.645858, -2.798684, -1.267847, 1.570796, 1.814192],accel_mss,speed_ms,0,blend_radius_m)
  movel([0.242724, -0.649188, -2.798339, -1.264862, 1.570796, 1.813520],accel_mss,speed_ms,0,blend_radius_m)
  movel([0.241608, -0.652588, -2.797982, -1.261820, 1.570796, 1.812404],accel_mss,speed_ms,0,blend_radius_m)
  movel([0.240439, -0.655954, -2.797623, -1.258811, 1.570796, 1.811236],accel_mss,speed_ms,0,blend_radius_m)
  movel([0.239603, -0.659200, -2.797273, -1.255916, 1.570796, 1.810399],accel_mss,speed_ms,0,blend_radius_m)
  movel([0.238338, -0.658028, -2.797400, -1.256960, 1.570796, 1.809135],accel_mss,speed_ms,0,blend_radius_m)
  movel([0.236551, -0.657567, -2.797450, -1.257372, 1.570796, 1.807347],accel_mss,speed_ms,0,blend_radius_m)
  movel([0.234295, -0.657870, -2.797417, -1.257101, 1.570796, 1.805091],accel_mss,speed_ms,0,blend_radius_m)
  movel([0.231615, -0.658998, -2.797295, -1.256096, 1.570796, 1.802411],accel_mss,speed_ms,0,blend_radius_m)
  speed_ms = 0.005
  movel([0.231615, -0.653180, -2.790577, -1.268632, 1.570796, 1.802411],accel_mss,speed_ms,0,blend_radius_m)
  speed_ms = 0.040
  movel([0.234282, -0.660908, -2.789729, -1.261752, 1.570796, 1.805079],accel_mss,speed_ms,0,blend_radius_m)
  speed_ms = 0.005
  movel([0.234282, -0.666838, -2.796431, -1.249120, 1.570796, 1.805079],accel_mss,speed_ms,0,blend_radius_m)
  speed_ms = 0.025
  movel([0.234647, -0.670305, -2.796040, -1.246043, 1.570796, 1.805443],accel_mss,speed_ms,0,blend_radius_m)
  movel([0.235625, -0.673194, -2.795711, -1.243484, 1.570796, 1.806421],accel_mss,speed_ms,0,blend_radius_m)
  movel([0.237414, -0.675104, -2.795491, -1.241794, 1.570796, 1.808211],accel_mss,speed_ms,0,blend_radius_m)
  movel([0.238680, -0.675565, -2.795438, -1.241387, 1.570796, 1.809476],accel_mss,speed_ms,0,blend_radius_m)
  movel([0.240229, -0.675630, -2.795430, -1.241329, 1.570796, 1.811025],accel_mss,speed_ms,0,blend_radius_m)
  movel([0.242736, -0.675031, -2.795500, -1.241858, 1.570796, 1.813533],accel_mss,speed_ms,0,blend_radius_m)
  movel([0.245485, -0.673775, -2.795644, -1.242970, 1.570796, 1.816282],accel_mss,speed_ms,0,blend_radius_m)
  movel([0.248430, -0.672010, -2.795847, -1.244533, 1.570796, 1.819227],accel_mss,speed_ms,0,blend_radius_m)
  movel([0.251520, -0.669886, -2.796088, -1.246415, 1.570796, 1.822316],accel_mss,speed_ms,0,blend_radius_m)
  movel([0.257922, -0.665161, -2.796618, -1.250610, 1.570796, 1.828718],accel_mss,speed_ms,0,blend_radius_m)
  movel([0.264253, -0.660832, -2.797095, -1.254462, 1.570796, 1.835049],accel_mss,speed_ms,0,blend_radius_m)
  movel([0.267743, -0.658968, -2.797298, -1.256122, 1.570796, 1.838540],accel_mss,speed_ms,0,blend_radius_m)
  movel([0.271017, -0.657713, -2.797434, -1.257241, 1.570796, 1.841814],accel_mss,speed_ms,0,blend_radius_m)
  movel([0.274016, -0.657063, -2.797504, -1.257821, 1.570796, 1.844813],accel_mss,speed_ms,0,blend_radius_m)
  movel([0.276680, -0.657024, -2.797508, -1.257856, 1.570796, 1.847476],accel_mss,speed_ms,0,blend_radius_m)
  movel([0.278959, -0.657579, -2.797449, -1.257362, 1.570796, 1.849755],accel_mss,speed_ms,0,blend_radius_m)
  movel([0.280797, -0.658728, -2.797324, -1.256337, 1.570796, 1.851594],accel_mss,speed_ms,0,blend_radius_m)
  movel([0.282138, -0.660462, -2.797136, -1.254791, 1.570796, 1.852934],accel_mss,speed_ms,0,blend_radius_m)
  movel([0.282941, -0.662761, -2.796884, -1.252745, 1.570796, 1.853738],accel_mss,speed_ms,0,blend_radius_m)
  speed_ms = 0.005
  movel([0.282941, -0.656889, -2.790174, -1.265327, 1.570796, 1.853738],accel_mss,speed_ms,0,blend_radius_m)
  speed_ms = 0.040
  movel([0.223582, -0.638749, -2.792092, -1.281548, 1.570796, 1.794378],accel_mss,speed_ms,0,blend_radius_m)
  speed_ms = 0.005
  movel([0.223582, -0.644352, -2.798838, -1.269198, 1.570796, 1.794378],accel_mss,speed_ms,0,blend_radius_m)
  speed_ms = 0.025
  movel([0.225135, -0.644371, -2.798836, -1.269181, 1.570796, 1.795931],accel_mss,speed_ms,0,blend_radius_m)
  movel([0.226263, -0.644971, -2.798775, -1.268643, 1.570796, 1.797059],accel_mss,speed_ms,0,blend_radius_m)
  movel([0.226487, -0.645669, -2.798703, -1.268017, 1.570796, 1.797283],accel_mss,speed_ms,0,blend_radius_m)
  movel([0.226392, -0.646641, -2.798603, -1.267145, 1.570796, 1.797188],accel_mss,speed_ms,0,blend_radius_m)
  movel([0.225968, -0.647782, -2.798485, -1.266122, 1.570796, 1.796765],accel_mss,speed_ms,0,blend_radius_m)
  movel([0.225199, -0.648989, -2.798360, -1.265041, 1.570796, 1.795995],accel_mss,speed_ms,0,blend_radius_m)
  movel([0.223413, -0.651070, -2.798142, -1.263177, 1.570796, 1.794209],accel_mss,speed_ms,0,blend_radius_m)
  movel([0.222779, -0.652196, -2.798023, -1.262169, 1.570796, 1.793575],accel_mss,speed_ms,0,blend_radius_m)
  movel([0.222508, -0.653206, -2.797916, -1.261266, 1.570796, 1.793304],accel_mss,speed_ms,0,blend_radius_m)
  movel([0.222726, -0.654769, -2.797750, -1.259870, 1.570796, 1.793522],accel_mss,speed_ms,0,blend_radius_m)
  movel([0.223558, -0.656028, -2.797615, -1.258745, 1.570796, 1.794355],accel_mss,speed_ms,0,blend_radius_m)
  movel([0.224721, -0.656896, -2.797522, -1.257971, 1.570796, 1.795518],accel_mss,speed_ms,0,blend_radius_m)
  movel([0.226187, -0.657371, -2.797471, -1.257547, 1.570796, 1.796983],accel_mss,speed_ms,0,blend_radius_m)
  movel([0.227923, -0.657433, -2.797464, -1.257491, 1.570796, 1.798720],accel_mss,speed_ms,0,blend_radius_m)
  movel([0.226480, -0.659962, -2.797190, -1.255236, 1.570796, 1.797277],accel_mss,speed_ms,0,blend_radius_m)
  movel([0.225397, -0.662372, -2.796927, -1.253090, 1.570796, 1.796193],accel_mss,speed_ms,0,blend_radius_m)
  movel([0.224628, -0.664667, -2.796673, -1.251049, 1.570796, 1.795424],accel_mss,speed_ms,0,blend_radius_m)
  movel([0.224130, -0.666844, -2.796430, -1.249114, 1.570796, 1.794927],accel_mss,speed_ms,0,blend_radius_m)
  movel([0.223789, -0.670845, -2.795979, -1.245565, 1.570796, 1.794586],accel_mss,speed_ms,0,blend_radius_m)
  movel([0.224067, -0.674358, -2.795577, -1.242454, 1.570796, 1.794863],accel_mss,speed_ms,0,blend_radius_m)
  movel([0.224409, -0.677690, -2.795191, -1.239508, 1.570796, 1.795206],accel_mss,speed_ms,0,blend_radius_m)
  movel([0.224276, -0.679569, -2.794971, -1.237849, 1.570796, 1.795072],accel_mss,speed_ms,0,blend_radius_m)
  movel([0.223747, -0.681697, -2.794720, -1.235972, 1.570796, 1.794543],accel_mss,speed_ms,0,blend_radius_m)
  movel([0.222635, -0.684121, -2.794431, -1.233837, 1.570796, 1.793431],accel_mss,speed_ms,0,blend_radius_m)
  movel([0.221002, -0.686579, -2.794136, -1.231673, 1.570796, 1.791799],accel_mss,speed_ms,0,blend_radius_m)
  movel([0.219067, -0.688694, -2.793880, -1.229815, 1.570796, 1.789863],accel_mss,speed_ms,0,blend_radius_m)
  movel([0.217059, -0.690075, -2.793712, -1.228602, 1.570796, 1.787855],accel_mss,speed_ms,0,blend_radius_m)
  movel([0.217832, -0.691093, -2.793587, -1.227709, 1.570796, 1.788628],accel_mss,speed_ms,0,blend_radius_m)
  movel([0.218587, -0.693931, -2.793237, -1.225221, 1.570796, 1.789383],accel_mss,speed_ms,0,blend_radius_m)
  movel([0.218569, -0.695692, -2.793018, -1.223679, 1.570796, 1.789365],accel_mss,speed_ms,0,blend_radius_m)
  movel([0.217778, -0.699726, -2.792511, -1.220152, 1.570796, 1.788574],accel_mss,speed_ms,0,blend_radius_m)
  movel([0.217007, -0.701936, -2.792230, -1.218223, 1.570796, 1.787803],accel_mss,speed_ms,0,blend_radius_m)
  movel([0.215989, -0.704239, -2.791935, -1.216215, 1.570796, 1.786785],accel_mss,speed_ms,0,blend_radius_m)
  speed_ms = 0.005
  movel([0.215989, -0.697796, -2.785314, -1.229278, 1.570796, 1.786785],accel_mss,speed_ms,0,blend_radius_m)
  speed_ms = 0.040
  movel([0.206248, -0.702773, -2.784671, -1.224945, 1.570796, 1.777044],accel_mss,speed_ms,0,blend_radius_m)
  speed_ms = 0.005
  movel([0.206248, -0.709281, -2.791281, -1.211827, 1.570796, 1.777044],accel_mss,speed_ms,0,blend_radius_m)
  speed_ms = 0.025
  movel([0.211186, -0.723264, -2.789404, -1.199721, 1.570796, 1.781982],accel_mss,speed_ms,0,blend_radius_m)
  movel([0.211525, -0.725206, -2.789136, -1.198047, 1.570796, 1.782322],accel_mss,speed_ms,0,blend_radius_m)
  movel([0.211317, -0.726404, -2.788970, -1.197015, 1.570796, 1.782113],accel_mss,speed_ms,0,blend_radius_m)
  movel([0.210680, -0.727770, -2.788780, -1.195840, 1.570796, 1.781476],accel_mss,speed_ms,0,blend_radius_m)
  movel([0.208591, -0.730766, -2.788359, -1.193264, 1.570796, 1.779387],accel_mss,speed_ms,0,blend_radius_m)
  movel([0.208183, -0.732155, -2.788163, -1.192071, 1.570796, 1.778979],accel_mss,speed_ms,0,blend_radius_m)
  movel([0.208317, -0.733223, -2.788011, -1.191155, 1.570796, 1.779114],accel_mss,speed_ms,0,blend_radius_m)
  movel([0.209180, -0.734404, -2.787843, -1.190143, 1.570796, 1.779976],accel_mss,speed_ms,0,blend_radius_m)
  movel([0.210570, -0.735048, -2.787751, -1.189591, 1.570796, 1.781366],accel_mss,speed_ms,0,blend_radius_m)
  movel([0.213649, -0.735829, -2.787639, -1.188921, 1.570796, 1.784445],accel_mss,speed_ms,0,blend_radius_m)
  movel([0.215273, -0.736891, -2.787486, -1.188012, 1.570796, 1.786069],accel_mss,speed_ms,0,blend_radius_m)
  movel([0.217074, -0.738970, -2.787186, -1.186233, 1.570796, 1.787870],accel_mss,speed_ms,0,blend_radius_m)
  movel([0.217550, -0.740234, -2.787002, -1.185153, 1.570796, 1.788347],accel_mss,speed_ms,0,blend_radius_m)
  movel([0.217501, -0.741551, -2.786810, -1.184029, 1.570796, 1.788298],accel_mss,speed_ms,0,blend_radius_m)
  movel([0.217217, -0.742207, -2.786714, -1.183468, 1.570796, 1.788013],accel_mss,speed_ms,0,blend_radius_m)
  movel([0.216727, -0.742851, -2.786619, -1.182919, 1.570796, 1.787523],accel_mss,speed_ms,0,blend_radius_m)
  movel([0.215036, -0.744079, -2.786438, -1.181872, 1.570796, 1.785832],accel_mss,speed_ms,0,blend_radius_m)
  movel([0.215175, -0.745359, -2.786249, -1.180780, 1.570796, 1.785971],accel_mss,speed_ms,0,blend_radius_m)
  movel([0.215769, -0.746452, -2.786087, -1.179850, 1.570796, 1.786565],accel_mss,speed_ms,0,blend_radius_m)
  movel([0.217876, -0.748132, -2.785837, -1.178420, 1.570796, 1.788672],accel_mss,speed_ms,0,blend_radius_m)
  movel([0.222717, -0.749972, -2.785561, -1.176856, 1.570796, 1.793513],accel_mss,speed_ms,0,blend_radius_m)
  movel([0.225551, -0.750262, -2.785517, -1.176610, 1.570796, 1.796347],accel_mss,speed_ms,0,blend_radius_m)
  movel([0.228744, -0.750201, -2.785526, -1.176661, 1.570796, 1.799541],accel_mss,speed_ms,0,blend_radius_m)
  movel([0.231573, -0.750614, -2.785464, -1.176311, 1.570796, 1.802369],accel_mss,speed_ms,0,blend_radius_m)
  movel([0.232625, -0.751249, -2.785368, -1.175771, 1.570796, 1.803421],accel_mss,speed_ms,0,blend_radius_m)
  movel([0.233314, -0.752306, -2.785209, -1.174875, 1.570796, 1.804110],accel_mss,speed_ms,0,blend_radius_m)
  movel([0.233415, -0.753093, -2.785089, -1.174207, 1.570796, 1.804211],accel_mss,speed_ms,0,blend_radius_m)
  movel([0.233239, -0.754071, -2.784940, -1.173377, 1.570796, 1.804035],accel_mss,speed_ms,0,blend_radius_m)
  movel([0.232768, -0.755072, -2.784787, -1.172529, 1.570796, 1.803564],accel_mss,speed_ms,0,blend_radius_m)
  movel([0.231974, -0.755926, -2.784657, -1.171806, 1.570796, 1.802771],accel_mss,speed_ms,0,blend_radius_m)
  movel([0.230645, -0.756409, -2.784583, -1.171397, 1.570796, 1.801441],accel_mss,speed_ms,0,blend_radius_m)
  movel([0.225181, -0.756582, -2.784556, -1.171251, 1.570796, 1.795978],accel_mss,speed_ms,0,blend_radius_m)
  movel([0.220271, -0.755833, -2.784671, -1.171885, 1.570796, 1.791068],accel_mss,speed_ms,0,blend_radius_m)
  movel([0.219820, -0.756948, -2.784500, -1.170941, 1.570796, 1.790616],accel_mss,speed_ms,0,blend_radius_m)
  movel([0.219625, -0.757947, -2.784346, -1.170096, 1.570796, 1.790421],accel_mss,speed_ms,0,blend_radius_m)
  movel([0.219903, -0.759619, -2.784087, -1.168683, 1.570796, 1.790699],accel_mss,speed_ms,0,blend_radius_m)
  movel([0.220890, -0.760902, -2.783888, -1.167599, 1.570796, 1.791686],accel_mss,speed_ms,0,blend_radius_m)
  movel([0.222361, -0.761874, -2.783736, -1.166779, 1.570796, 1.793158],accel_mss,speed_ms,0,blend_radius_m)
  movel([0.225953, -0.763076, -2.783548, -1.165765, 1.570796, 1.796749],accel_mss,speed_ms,0,blend_radius_m)
  movel([0.229001, -0.763673, -2.783454, -1.165262, 1.570796, 1.799798],accel_mss,speed_ms,0,blend_radius_m)
  movel([0.230012, -0.764065, -2.783393, -1.164932, 1.570796, 1.800808],accel_mss,speed_ms,0,blend_radius_m)
  movel([0.230275, -0.764506, -2.783323, -1.164560, 1.570796, 1.801072],accel_mss,speed_ms,0,blend_radius_m)
  movel([0.230233, -0.765201, -2.783213, -1.163975, 1.570796, 1.801029],accel_mss,speed_ms,0,blend_radius_m)
  movel([0.229847, -0.766112, -2.783069, -1.163208, 1.570796, 1.800643],accel_mss,speed_ms,0,blend_radius_m)
  movel([0.229315, -0.766807, -2.782959, -1.162623, 1.570796, 1.800112],accel_mss,speed_ms,0,blend_radius_m)
  movel([0.227997, -0.767766, -2.782807, -1.161816, 1.570796, 1.798794],accel_mss,speed_ms,0,blend_radius_m)
  movel([0.226146, -0.768931, -2.782621, -1.160837, 1.570796, 1.796942],accel_mss,speed_ms,0,blend_radius_m)
  movel([0.225764, -0.769458, -2.782537, -1.160395, 1.570796, 1.796561],accel_mss,speed_ms,0,blend_radius_m)
  movel([0.225546, -0.770196, -2.782418, -1.159774, 1.570796, 1.796343],accel_mss,speed_ms,0,blend_radius_m)
  movel([0.225620, -0.770833, -2.782316, -1.159240, 1.570796, 1.796416],accel_mss,speed_ms,0,blend_radius_m)
  movel([0.226374, -0.771831, -2.782155, -1.158403, 1.570796, 1.797170],accel_mss,speed_ms,0,blend_radius_m)
  movel([0.228390, -0.773025, -2.781962, -1.157402, 1.570796, 1.799186],accel_mss,speed_ms,0,blend_radius_m)
  movel([0.237740, -0.777024, -2.781311, -1.154054, 1.570796, 1.808536],accel_mss,speed_ms,0,blend_radius_m)
